(* IEC 61131-3 sources: JingjiangMoonbox/Application/Application/任务列表/Main_Task/IO列表 (part 2) *)

(* ---- KS_FB_MapAxisIOExtra.st ---- *)
(*@CES
Name=KS_FB_MapAxisIOExtra
Type=FunctionBlock
TypeGuid=6f9dac99-8de1-4efc-8465-68ac443b7d08
Guid=6be90e54-b934-4bee-925a-ddca26256504
HasDeclaration=True
HasImplementation=True
*)
{DECLARATION}
FUNCTION_BLOCK KS_FB_MapAxisIOExtra
VAR_INPUT
	i_xEn									: BOOL;(*功能块使能|*)
	i_xEnableInput							: BOOL;(*使能输入|*)
	i_xEnableOutput							: BOOL;(*使能输出|*)
	i_pstStIOMap_Axis_Extra_FE			: POINTER TO StIOMap_Axis_Extra_FE;(*轴io数据区域|*)

	i_xPreHeating							: BOOL; (* 预加热 *)
	i_xPreHeating_Err						: BOOL; (* 预加热报警\温控信号 *)
	i_xPreHotBlower							: BOOL; (* 预热风 *)
	i_xPreHotBlower_Err						: BOOL; (* 预热风报警 *)
	i_xCoolBlower							: BOOL; (* 冷风开关 *)
	i_xCoolBlower_Button					: BOOL; (* 冷风按钮 *)
	i_xCoolBlower_Err						: BOOL; (* 冷风报警 *)
	i_xHotBlower							: BOOL; (* 热风开关 *)
	i_xHotBlower_Button						: BOOL; (* 热风按钮 *)
	i_xHotBlower_Err						: BOOL; (* 热风报警 *)
	i_xHotBlower_Opened_Act					: BOOL; (* 热风实际被打开了|2022.5.11.192858|没有反馈时候需要写true*)
	i_xHotBlower_CHNL2						: BOOL; (* 第2路热风开关 *)
	i_xHotBlower_Button_CHNL2				: BOOL; (* 第2路热风按钮 *)
	i_xHotBlower_Err_CHNL2					: BOOL; (* 第2路热风报警 *)
	i_xHotBlower_Opened_Act_CHNL2			: BOOL; (* 热风2实际被打开了|2022.5.11.192858|没有反馈时候需要写true*)
	i_xTemReachToTarget						: BOOL; (* 到达目标温度 *)
	i_xSteamHeating							: BOOL; (* 蒸汽加热开关 *)
	i_xSteamHeating_Err						: BOOL; (* 蒸汽加热报警 *)
	i_xHeating_I							: BOOL; (* 电加热I档 *)
	i_xHeating_II							: BOOL; (* 电加热II档 *)
	i_xHeating_III							: BOOL; (* 电加热III档 *)
	i_xHeating_Button						: BOOL; (* 加热按钮 *)
	i_xHeating_I_CHNL2						: BOOL; (* 第2路电加热I档 *)
	i_xHeating_II_CHNL2						: BOOL; (* 第2路电加热II档 *)
	i_xHeating_III_CHNL2					: BOOL; (* 第2路电加热III档 *)
	i_xHeating_Button_CHNL2					: BOOL; (* 第2路加热按钮 *)
	i_xAllExhBlower_Up						: BOOL; (* 全上排风 *)
	i_xAllExhBlower_Err_Up					: BOOL; (* 上排风报警 *)
	i_xAllExhBlower_Dn						: BOOL; (* 全下排风 *)
	i_xAllExhBlower_Err_Dn					: BOOL; (* 下排风报警 *)
	i_xAllCoolBlower						: BOOL; (* 全冷风 *)
	i_xAllHotBlower							: BOOL; (* 全热风 *)
	i_xAllHeating							: BOOL; (* 全加热 *)
	i_xAirInletMotorMin_Limit				: BOOL; (* 进风口风门电机最小开度限位 *)
	i_xAirInletMotorMax_Limit				: BOOL; (* 进风口风门电机最大开度限位 *)
	i_xOvensAirOutMotorMin_Limit			: BOOL; (* 烘箱出风口风门电机最小开度限位 *)
	i_xOvensAirOutMotorMax_Limit			: BOOL; (* 烘箱出风口风门电机最大开度限位 *)
	i_xAirExhaustMotorMin_Limit				: BOOL; (* 排风口风门电机最小开度限位 *)
	i_xAirExhaustMotorMax_Limit				: BOOL; (* 排风口风门电机最大开度限位 *)
	i_xAirReturnMotorMin_Limit				: BOOL; (* 回风口风门电机最小开度限位 *)
	i_xAirReturnMotorMax_Limit				: BOOL; (* 回风口风门电机最大开度限位 *)
	i_xScraperInveterError					: BOOL; (* 刮刀变频器报警 *)
	i_xScraperOn							: BOOL; (* 刮刀开关 *)
	i_xInkRollerInveterError				: BOOL; (* 递墨辊变频器报警 |2022.3.26.094940*)
	i_xInkRoller_CW							: BOOL; (* 递墨辊正转开 *)
	i_xInkRoller_CCW						: BOOL; (* 递墨辊反转开 *)
	i_xInkRoller_Up							: BOOL; (* 递墨辊上 *)
	i_xInkRoller_Dn							: BOOL; (* 递墨辊下 *)
	i_xTurnoverFilmAgency					: BOOL; (* 翻料架开关 *)
	i_wAI_AirInletMotor						: WORD; (* 进风口反馈|模拟量控制风门LEL *)
	i_wAI_OvensAirOutMotor					: WORD; (* 烘箱出风口反馈|模拟量控制风门LEL *)
	i_wAI_AirExhaustMotor					: WORD; (* 排风口反馈|模拟量控制风门LEL *)
	i_wAI_AirReturnMotor					: WORD; (* 回风反馈|模拟量控制风门LEL *)
	i_wInputLel								: WORD; (* LEL浓度反馈 *)
	i_wInAllAir								: WORD; (* 总进风反馈输入 *)
	i_wInFreshAir							: WORD; (* 新风反馈输入 *)
	i_wInExhaustAir							: WORD; (* 排风反馈输入 *)
	i_wInReturnAir							: WORD; (* 二次回风反馈输入 *)
	i_xTaper_Incr							: BOOL; (* 增加锥度+|针对牵引 *)
	i_xTaper_Decr							: BOOL; (* 减小锥度-|针对牵引 *)
	i_wAI_CoatingSensor						: WORD; (* 涂布传感器模拟量 *)
	i_byAIType_CoatingSensor				: BYTE; (* 涂布传感器类型 *)
	i_xAirExhaustSwitch						: BOOL; (* 色组排风输入开关 *)
	i_xAirExhaustButton						: BOOL; (* 色组排风输入按钮 *)
	i_xPushIn_PrnRoller						: BOOL; (* 顶版-进 *)
	i_xPullOut_PrnRoller					: BOOL; (* 顶版-退 *)
	i_xRsvd_DI0								: BOOL; (* 数字量输入保留0 *)
	i_xRsvd_DI1								: BOOL; (* 数字量输入保留1 *)
	i_xRsvd_DI2								: BOOL; (* 数字量输入保留2 *)
	i_xRsvd_DI3								: BOOL; (* 数字量输入保留3 *)
	i_xRsvd_DI4								: BOOL; (* 数字量输入保留4 *)
	i_xRsvd_DI5								: BOOL; (* 数字量输入保留5 *)
	i_xRsvd_DI6								: BOOL; (* 数字量输入保留6 *)
	i_xRsvd_DI7								: BOOL; (* 数字量输入保留7 *)
	i_xRsvd_DI8								: BOOL; (* 数字量输入保留8 *)
	i_xRsvd_DI9								: BOOL; (* 数字量输入保留9 *)
	i_xRsvd_DI10							: BOOL; (* 数字量输入保留10 *)
	i_xRsvd_DI11							: BOOL; (* 数字量输入保留11 *)
	i_xRsvd_DI12							: BOOL; (* 数字量输入保留12 *)
	i_xRsvd_DI13							: BOOL; (* 数字量输入保留13 *)
	i_xRsvd_DI14							: BOOL; (* 数字量输入保留14 *)
	i_xRsvd_DI15							: BOOL; (* 数字量输入保留15 *)
	i_wRsvd_AI0								: WORD; (* 模拟量输入保留0 *)
	i_wRsvd_AI1								: WORD; (* 模拟量输入保留1 *)
	i_wRsvd_AI2								: WORD; (* 模拟量输入保留2 *)
	i_wRsvd_AI3								: WORD; (* 模拟量输入保留3 *)
	i_wRsvd_AI4								: WORD; (* 模拟量输入保留4 *)
	i_wRsvd_AI5								: WORD; (* 模拟量输入保留5 *)

END_VAR
VAR_OUTPUT
	o_xEno									: BOOL;
	o_iErNo									: INT;

	o_xRel_PreHeating						: BOOL; (* 预加热接触器 *)
	o_xLamp_PreHeating						: BOOL; (* 预加热指示灯 *)
	o_xRel_ResetErr_PreHeating				: BOOL; (* 预加热故障复位 *)
	o_wAO_PreHeating						: WORD; (* 预加热模拟量 *)
	o_xRel_PreHeatingRoller_Motor			: BOOL; (* 预热辊使能 *)
	o_xRel_PreHeatingRoller_Motor_Rev		: BOOL; (* 预热辊反转使能 *)
	o_wAO_PreHeatingRoller_Motor			: WORD; (* 预热辊模拟量输出 *)
	o_xRel_PreHotBlower						: BOOL; (* 预热风接触器 *)
	o_xLamp_PreHotBlower					: BOOL; (* 预热风指示灯 *)
	o_xRel_ResetErr_PreHotBlower			: BOOL; (* 预热风故障复位 *)
	o_wAO_PreHotBlower						: WORD; (* 预热风模拟量 *)
	o_xRel_CoolBlower						: BOOL; (* 冷风接触器 *)
	o_xLamp_CoolBlower						: BOOL; (* 冷风指示灯 *)
	o_xRel_HotBlower						: BOOL; (* 热风接触器 *)
	o_xLamp_HotBlower						: BOOL; (* 热风指示灯 *)
	o_xRel_ResetErr_HotBlower				: BOOL; (* 热风故障复位 *)
	o_wAO_HotBlower							: WORD; (* 热风模拟量输出 *)
	o_xRel_HotBlower_CHNL2					: BOOL; (* 第2路热风接触器 *)
	o_xLamp_HotBlower_CHNL2					: BOOL; (* 第2路热风指示灯 *)
	o_xRel_ResetErr_HotBlower_CHNL2			: BOOL; (* 第2路热风故障复位 *)
	o_wAO_HotBlower_CHNL2					: WORD; (* 第2路热风模拟量输出 *)
	o_xRel_SteamHeating						: BOOL; (* 蒸汽输出 *)
	o_xLamp_SteamHeating					: BOOL; (* 蒸汽加热指示灯 *)
	o_xRel_ResetErr_SteamHeating			: BOOL; (* 蒸汽加热复位 *)
	o_wAO_SteamHeating						: WORD; (* 蒸汽加热模拟量输出 *)
	o_xRel_Heating_I						: BOOL; (* 电加热I档 *)
	o_xRel_Heating_II						: BOOL; (* 电加热II档 *)
	o_xRel_Heating_III						: BOOL; (* 电加热III档 *)
	o_xLamp_Heating							: BOOL; (* 电加热指示灯 *)
	o_xRel_Heating_I_CHNL2					: BOOL; (* 第2路电加热I档 *)
	o_xRel_Heating_II_CHNL2					: BOOL; (* 第2路电加热II档 *)
	o_xRel_Heating_III_CHNL2				: BOOL; (* 第2路电加热III档 *)
	o_xLamp_Heating_CHNL2					: BOOL; (* 第2路电加热指示灯 *)
	o_xRel_AllExhBlower_Up					: BOOL; (* 上排风继电器输出 *)
	o_xLamp_AllExhBlower_Up					: BOOL; (* 全上排风指示灯 *)
	o_xRel_ModeStar_AllExhBlower_Up			: BOOL; (* 上排风模式-星形 *)
	o_xRel_ModeTriangle_AllExhBlower_Up		: BOOL; (* 上排风模式-三角 *)
	o_xRel_ResetErr_AllExhBlower_Up			: BOOL; (* 上排风故障复位 *)
	o_wAO_AllExhBlower_Up					: WORD; (* 上排风模拟量输出 *)
	o_xRel_AllExhBlower_Dn					: BOOL; (* 下排风继电器输出 *)
	o_xLamp_AllExhBlower_Dn					: BOOL; (* 全下排风指示灯 *)
	o_xRel_ModeStar_AllExhBlower_Dn			: BOOL; (* 下排风模式-星形 *)
	o_xRel_ModeTriangle_AllExhBlower_Dn		: BOOL; (* 下排风模式-三角 *)
	o_xRel_ResetErr_AllExhBlower_Dn			: BOOL; (* 下排风故障复位 *)
	o_wAO_AllExhBlower_Dn					: WORD; (* 下排风模拟量输出 *)
	o_xLamp_AllCoolBlower					: BOOL; (* 全冷风指示灯 *)
	o_xLamp_AllHotBlower					: BOOL; (* 全热风指示灯 *)
	o_xLamp_AllHeating						: BOOL; (* 全加热指示灯 *)
	o_xAirInletMotor_Increase				: BOOL; (* 进风口风门开度增大 *)
	o_xAirInletMotor_Decrease				: BOOL; (* 进风口风门开度减小 *)
	o_xOvensAirOutMotor_Increase			: BOOL; (* 烘箱出风口风门开度增大 *)
	o_xOvensAirOutMotor_Decrease			: BOOL; (* 烘箱出风口风门开度减小 *)
	o_xAirExhaustMotor_Increase				: BOOL; (* 排风口风门开度增大 *)
	o_xAirExhaustMotor_Decrease				: BOOL; (* 排风口风门开度减小 *)
	o_xAirReturnMotor_Increase				: BOOL; (* 回风风门开度增大 *)
	o_xAirReturnMotor_Decrease				: BOOL; (* 回风风门开度减小 *)
	o_xScraperOn							: BOOL; (* 刮刀输出 *)
	o_xScraperRst							: BOOL;(*刮刀故障复位*)
	o_wAO_Scraper							: WORD; (* 刮刀模拟量输出 *)
	o_xInkRollerOn							: BOOL; (* 递墨辊运动信号 *)
	o_xInkRollerRst							: BOOL;(*递墨辊复位2022.7.8.093223*)
	o_xRel_InkRoller_CW						: BOOL; (* 递墨辊正转 *)
	o_xRel_InkRoller_CCW					: BOOL; (* 递墨辊反转 *)
	o_wAO_InkRoller							: WORD; (* 递墨辊模拟量输出 *)
	(*2026.05.25.135151*)
	o_wAO_InkRoller_Dir						: WORD;(* 递墨辊模拟量输出@±10V *)
	o_xRel_InkRoller_Up						: BOOL; (* 递墨辊上输出 *)
	o_xRel_InkRoller_Dn						: BOOL; (* 递墨辊下输出 *)
	o_xRel_TurnoverFilmAgency				: BOOL; (* 翻料架输出 *)
	o_xRel_ColdWaterRoller_Motor			: BOOL; (* 水冷辊电机使能 *)
	o_xRel_ColdWaterRoller_Motor_Rev		: BOOL; (* 水冷辊电机反转使能 *)
	o_wAO_ColdWaterRoller_Motor				: WORD; (* 水冷辊电机模拟量输出 *)
	o_xRel_DriveAfterPrint_Motor			: BOOL; (* 印后传动辊电机使能 *)
	o_xRel_DriveAfterPrint_Motor_Rev		: BOOL; (* 印后传动辊电机反转 *)
	o_wAO_DriveAfterPrint_Motor				: WORD; (* 印后传动辊电机模拟量输出 *)
	o_wAO_AirInletMotor						: WORD; (* 进口输出|模拟量控制风门LEL *)
	o_wAO_OvensAirOutMotor					: WORD; (* 烘箱出风口输出|模拟量控制风门LEL *)
	o_wAO_AirExhaustMotor					: WORD; (* 排风口输出|模拟量控制风门LEL *)
	o_wAO_AirReturnMotor					: WORD; (* 回风输出|模拟量控制风门LEL *)
	o_wInAllAir								: WORD; (* 总进风输出 *)
	o_wInFreshAir							: WORD; (* 新风输出 *)
	o_wInExhaustAir							: WORD; (* 排风输出 *)
	o_wInReturnAir							: WORD; (* 二次回风输出 *)
	o_wPreAirHotRollTorque					: WORD; (* 预热辊转矩输出 *)
	o_wCoolWaterRollTorque					: WORD; (* 水冷辊转矩输出 *)
	o_xAirExhaustEn							: BOOL; (* 色组排风输出使能 *)
	o_xRel_PushIn_PrnRoller					: BOOL; (* 顶版-进执行 *)
	o_xRel_PullOut_PrnRoller				: BOOL; (* 顶版-退执行 *)
	o_xRel_ModeStar_HotBlower				: BOOL; (* 热风输出-星形 *)
	o_xRel_ModeTriangle_HotBlower			: BOOL; (* 热风输出-三角 *)
	o_xRel_Oven								: BOOL; (* 色组烘箱输出 *)
	o_xRsvd_DO0								: BOOL; (* 数字量输出保留0 *)
	o_xRsvd_DO1								: BOOL; (* 数字量输出保留1 *)
	o_xRsvd_DO2								: BOOL; (* 数字量输出保留2 *)
	o_xRsvd_DO3								: BOOL; (* 数字量输出保留3 *)
	o_xRsvd_DO4								: BOOL; (* 数字量输出保留4 *)
	o_xRsvd_DO5								: BOOL; (* 数字量输出保留5 *)
	o_xRsvd_DO6								: BOOL; (* 数字量输出保留6 *)
	o_xRsvd_DO7								: BOOL; (* 数字量输出保留7 *)
	o_xRsvd_DO8								: BOOL; (* 数字量输出保留8 *)
	o_xRsvd_DO9								: BOOL; (* 数字量输出保留9 *)
	o_xRsvd_DO10							: BOOL; (* 数字量输出保留10 *)
	o_xRsvd_DO11							: BOOL; (* 数字量输出保留11 *)
	o_xRsvd_DO12							: BOOL; (* 数字量输出保留12 *)
	o_xRsvd_DO13							: BOOL; (* 数字量输出保留13 *)
	o_xRsvd_DO14							: BOOL; (* 数字量输出保留14 *)
	o_xRsvd_DO15							: BOOL; (* 数字量输出保留15 *)
	o_wRsvd_AO0								: WORD; (* 模拟量输出保留0 *)
	o_wRsvd_AO1								: WORD; (* 模拟量输出保留1 *)
	o_wRsvd_AO2								: WORD; (* 模拟量输出保留2 *)
	o_wRsvd_AO3								: WORD; (* 模拟量输出保留3 *)
	o_wRsvd_AO4								: WORD; (* 模拟量输出保留4 *)
	o_wRsvd_AO5								: WORD; (* 模拟量输出保留5 *)
END_VAR
VAR
END_VAR

{IMPLEMENTATION}
o_xEno:= i_xEn;
o_iErNo:= 0;
IF i_xEn THEN
	IF i_pstStIOMap_Axis_Extra_FE<>0 THEN
		IF i_xEnableInput THEN (* 输入 *)
			i_pstStIOMap_Axis_Extra_FE^.i_xPreHeating					:= i_xPreHeating					;//		: BOOL; (* 预加热 *)
			i_pstStIOMap_Axis_Extra_FE^.i_xPreHeating_Err				:= i_xPreHeating_Err				;//		: BOOL; (* 预加热报警\温控信号 *)
			i_pstStIOMap_Axis_Extra_FE^.i_xPreHotBlower					:= i_xPreHotBlower					;//		: BOOL; (* 预热风 *)
			i_pstStIOMap_Axis_Extra_FE^.i_xPreHotBlower_Err				:= i_xPreHotBlower_Err				;//		: BOOL; (* 预热风报警 *)
			i_pstStIOMap_Axis_Extra_FE^.i_xCoolBlower					:= i_xCoolBlower					;//		: BOOL; (* 冷风开关 *)
			i_pstStIOMap_Axis_Extra_FE^.i_xCoolBlower_Button				:= i_xCoolBlower_Button				;//		: BOOL; (* 冷风按钮 *)
			i_pstStIOMap_Axis_Extra_FE^.i_xCoolBlower_Err				:= i_xCoolBlower_Err				;//		: BOOL; (* 冷风报警 *)
			i_pstStIOMap_Axis_Extra_FE^.i_xHotBlower						:= i_xHotBlower						;//		: BOOL; (* 热风开关 *)
			i_pstStIOMap_Axis_Extra_FE^.i_xHotBlower_Button				:= i_xHotBlower_Button				;//		: BOOL; (* 热风按钮 *)
			i_pstStIOMap_Axis_Extra_FE^.i_xHotBlower_Err					:= i_xHotBlower_Err					;//		: BOOL; (* 热风报警 *)
			i_pstStIOMap_Axis_Extra_FE^.i_xHotBlower_Opened_Act			:= i_xHotBlower_Opened_Act			;//		: BOOL; (* 热风实际被打开了|2022.5.11.192858|没有反馈时候需要写true*)
			i_pstStIOMap_Axis_Extra_FE^.i_xHotBlower_CHNL2				:= i_xHotBlower_CHNL2				;//		: BOOL; (* 第2路热风开关 *)
			i_pstStIOMap_Axis_Extra_FE^.i_xHotBlower_Button_CHNL2		:= i_xHotBlower_Button_CHNL2		;//		: BOOL; (* 第2路热风按钮 *)
			i_pstStIOMap_Axis_Extra_FE^.i_xHotBlower_Err_CHNL2			:= i_xHotBlower_Err_CHNL2			;//		: BOOL; (* 第2路热风报警 *)
			i_pstStIOMap_Axis_Extra_FE^.i_xHotBlower_Opened_Act_CHNL2	:= i_xHotBlower_Opened_Act_CHNL2	;//		: BOOL; (* 热风2实际被打开了|2022.5.11.192858|没有反馈时候需要写true*)
			i_pstStIOMap_Axis_Extra_FE^.i_xTemReachToTarget				:= i_xTemReachToTarget				;//		: BOOL; (* 到达目标温度 *)
			i_pstStIOMap_Axis_Extra_FE^.i_xSteamHeating					:= i_xSteamHeating					;//		: BOOL; (* 蒸汽加热开关 *)
			i_pstStIOMap_Axis_Extra_FE^.i_xSteamHeating_Err				:= i_xSteamHeating_Err				;//		: BOOL; (* 蒸汽加热报警 *)
			i_pstStIOMap_Axis_Extra_FE^.i_xHeating_I						:= i_xHeating_I						;//		: BOOL; (* 电加热I档 *)
			i_pstStIOMap_Axis_Extra_FE^.i_xHeating_II					:= i_xHeating_II					;//		: BOOL; (* 电加热II档 *)
			i_pstStIOMap_Axis_Extra_FE^.i_xHeating_III					:= i_xHeating_III					;//		: BOOL; (* 电加热III档 *)
			i_pstStIOMap_Axis_Extra_FE^.i_xHeating_Button				:= i_xHeating_Button				;//		: BOOL; (* 加热按钮 *)
			i_pstStIOMap_Axis_Extra_FE^.i_xHeating_I_CHNL2				:= i_xHeating_I_CHNL2				;//		: BOOL; (* 第2路电加热I档 *)
			i_pstStIOMap_Axis_Extra_FE^.i_xHeating_II_CHNL2				:= i_xHeating_II_CHNL2				;//		: BOOL; (* 第2路电加热II档 *)
			i_pstStIOMap_Axis_Extra_FE^.i_xHeating_III_CHNL2				:= i_xHeating_III_CHNL2				;//		: BOOL; (* 第2路电加热III档 *)
			i_pstStIOMap_Axis_Extra_FE^.i_xHeating_Button_CHNL2			:= i_xHeating_Button_CHNL2			;//		: BOOL; (* 第2路加热按钮 *)
			i_pstStIOMap_Axis_Extra_FE^.i_xAllExhBlower_Up				:= i_xAllExhBlower_Up				;//		: BOOL; (* 全上排风 *)
			i_pstStIOMap_Axis_Extra_FE^.i_xAllExhBlower_Err_Up			:= i_xAllExhBlower_Err_Up			;//		: BOOL; (* 上排风报警 *)
			i_pstStIOMap_Axis_Extra_FE^.i_xAllExhBlower_Dn				:= i_xAllExhBlower_Dn				;//		: BOOL; (* 全下排风 *)
			i_pstStIOMap_Axis_Extra_FE^.i_xAllExhBlower_Err_Dn			:= i_xAllExhBlower_Err_Dn			;//		: BOOL; (* 下排风报警 *)
			i_pstStIOMap_Axis_Extra_FE^.i_xAllCoolBlower					:= i_xAllCoolBlower					;//		: BOOL; (* 全冷风 *)
			i_pstStIOMap_Axis_Extra_FE^.i_xAllHotBlower					:= i_xAllHotBlower					;//		: BOOL; (* 全热风 *)
			i_pstStIOMap_Axis_Extra_FE^.i_xAllHeating					:= i_xAllHeating					;//		: BOOL; (* 全加热 *)
			i_pstStIOMap_Axis_Extra_FE^.i_xAirInletMotorMin_Limit		:= i_xAirInletMotorMin_Limit		;//		: BOOL; (* 进风口风门电机最小开度限位 *)
			i_pstStIOMap_Axis_Extra_FE^.i_xAirInletMotorMax_Limit		:= i_xAirInletMotorMax_Limit		;//		: BOOL; (* 进风口风门电机最大开度限位 *)
			i_pstStIOMap_Axis_Extra_FE^.i_xOvensAirOutMotorMin_Limit		:= i_xOvensAirOutMotorMin_Limit		;//		: BOOL; (* 烘箱出风口风门电机最小开度限位 *)
			i_pstStIOMap_Axis_Extra_FE^.i_xOvensAirOutMotorMax_Limit		:= i_xOvensAirOutMotorMax_Limit		;//		: BOOL; (* 烘箱出风口风门电机最大开度限位 *)
			i_pstStIOMap_Axis_Extra_FE^.i_xAirExhaustMotorMin_Limit		:= i_xAirExhaustMotorMin_Limit		;//		: BOOL; (* 排风口风门电机最小开度限位 *)
			i_pstStIOMap_Axis_Extra_FE^.i_xAirExhaustMotorMax_Limit		:= i_xAirExhaustMotorMax_Limit		;//		: BOOL; (* 排风口风门电机最大开度限位 *)
			i_pstStIOMap_Axis_Extra_FE^.i_xAirReturnMotorMin_Limit		:= i_xAirReturnMotorMin_Limit		;//		: BOOL; (* 回风口风门电机最小开度限位 *)
			i_pstStIOMap_Axis_Extra_FE^.i_xAirReturnMotorMax_Limit		:= i_xAirReturnMotorMax_Limit		;//		: BOOL; (* 回风口风门电机最大开度限位 *)
			i_pstStIOMap_Axis_Extra_FE^.i_xScraperInveterError			:= i_xScraperInveterError			;//		: BOOL; (* 刮刀变频器报警 *)
			i_pstStIOMap_Axis_Extra_FE^.i_xScraperOn						:= i_xScraperOn						;//		: BOOL; (* 刮刀开关 *)
			i_pstStIOMap_Axis_Extra_FE^.i_xInkRollerInveterError			:= i_xInkRollerInveterError			;//		: BOOL; (* 递墨辊变频器报警 |2022.3.26.094940*)
			i_pstStIOMap_Axis_Extra_FE^.i_xInkRoller_CW					:= i_xInkRoller_CW					;//		: BOOL; (* 递墨辊正转开 *)
			i_pstStIOMap_Axis_Extra_FE^.i_xInkRoller_CCW					:= i_xInkRoller_CCW					;//		: BOOL; (* 递墨辊反转开 *)
			i_pstStIOMap_Axis_Extra_FE^.i_xInkRoller_Up					:= i_xInkRoller_Up					;//		: BOOL; (* 递墨辊上 *)
			i_pstStIOMap_Axis_Extra_FE^.i_xInkRoller_Dn					:= i_xInkRoller_Dn					;//		: BOOL; (* 递墨辊下 *)
			i_pstStIOMap_Axis_Extra_FE^.i_xTurnoverFilmAgency			:= i_xTurnoverFilmAgency			;//		: BOOL; (* 翻料架开关 *)
			i_pstStIOMap_Axis_Extra_FE^.i_wAI_AirInletMotor				:= i_wAI_AirInletMotor				;//		: WORD; (* 进风口反馈|模拟量控制风门LEL *)
			i_pstStIOMap_Axis_Extra_FE^.i_wAI_OvensAirOutMotor			:= i_wAI_OvensAirOutMotor			;//		: WORD; (* 烘箱出风口反馈|模拟量控制风门LEL *)
			i_pstStIOMap_Axis_Extra_FE^.i_wAI_AirExhaustMotor			:= i_wAI_AirExhaustMotor			;//		: WORD; (* 排风口反馈|模拟量控制风门LEL *)
			i_pstStIOMap_Axis_Extra_FE^.i_wAI_AirReturnMotor				:= i_wAI_AirReturnMotor				;//		: WORD; (* 回风反馈|模拟量控制风门LEL *)
			i_pstStIOMap_Axis_Extra_FE^.i_wInputLel						:= i_wInputLel						;//		: WORD; (* LEL浓度反馈 *)
			i_pstStIOMap_Axis_Extra_FE^.i_wInAllAir						:= i_wInAllAir						;//		: WORD; (* 总进风反馈输入 *)
			i_pstStIOMap_Axis_Extra_FE^.i_wInFreshAir					:= i_wInFreshAir					;//		: WORD; (* 新风反馈输入 *)
			i_pstStIOMap_Axis_Extra_FE^.i_wInExhaustAir					:= i_wInExhaustAir					;//		: WORD; (* 排风反馈输入 *)
			i_pstStIOMap_Axis_Extra_FE^.i_wInReturnAir					:= i_wInReturnAir					;//		: WORD; (* 二次回风反馈输入 *)
			i_pstStIOMap_Axis_Extra_FE^.i_xTaper_Incr					:= i_xTaper_Incr					;//		: BOOL; (* 增加锥度+|针对牵引 *)
			i_pstStIOMap_Axis_Extra_FE^.i_xTaper_Decr					:= i_xTaper_Decr					;//		: BOOL; (* 减小锥度-|针对牵引 *)
			i_pstStIOMap_Axis_Extra_FE^.i_wAI_CoatingSensor				:= i_wAI_CoatingSensor				;//		: WORD; (* 涂布传感器模拟量 *)
			i_pstStIOMap_Axis_Extra_FE^.i_byAIType_CoatingSensor			:= i_byAIType_CoatingSensor			;//		: BYTE; (* 涂布传感器类型 *)
			i_pstStIOMap_Axis_Extra_FE^.i_xAirExhaustSwitch				:= i_xAirExhaustSwitch				;//		: BOOL; (* 色组排风输入开关 *)
			i_pstStIOMap_Axis_Extra_FE^.i_xAirExhaustButton				:= i_xAirExhaustButton				;//		: BOOL; (* 色组排风输入按钮 *)
			i_pstStIOMap_Axis_Extra_FE^.i_xPushIn_PrnRoller				:= i_xPushIn_PrnRoller				;//		: BOOL; (* 顶版-进 *)
			i_pstStIOMap_Axis_Extra_FE^.i_xPullOut_PrnRoller				:= i_xPullOut_PrnRoller				;//		: BOOL; (* 顶版-退 *)
			i_pstStIOMap_Axis_Extra_FE^.i_xRsvd_DI0						:= i_xRsvd_DI0						;//		: BOOL; (* 数字量输入保留0 *)
			i_pstStIOMap_Axis_Extra_FE^.i_xRsvd_DI1						:= i_xRsvd_DI1						;//		: BOOL; (* 数字量输入保留1 *)
			i_pstStIOMap_Axis_Extra_FE^.i_xRsvd_DI2						:= i_xRsvd_DI2						;//		: BOOL; (* 数字量输入保留2 *)
			i_pstStIOMap_Axis_Extra_FE^.i_xRsvd_DI3						:= i_xRsvd_DI3						;//		: BOOL; (* 数字量输入保留3 *)
			i_pstStIOMap_Axis_Extra_FE^.i_xRsvd_DI4						:= i_xRsvd_DI4						;//		: BOOL; (* 数字量输入保留4 *)
			i_pstStIOMap_Axis_Extra_FE^.i_xRsvd_DI5						:= i_xRsvd_DI5						;//		: BOOL; (* 数字量输入保留5 *)
			i_pstStIOMap_Axis_Extra_FE^.i_xRsvd_DI6						:= i_xRsvd_DI6						;//		: BOOL; (* 数字量输入保留6 *)
			i_pstStIOMap_Axis_Extra_FE^.i_xRsvd_DI7						:= i_xRsvd_DI7						;//		: BOOL; (* 数字量输入保留7 *)
			i_pstStIOMap_Axis_Extra_FE^.i_xRsvd_DI8						:= i_xRsvd_DI8						;//		: BOOL; (* 数字量输入保留8 *)
			i_pstStIOMap_Axis_Extra_FE^.i_xRsvd_DI9						:= i_xRsvd_DI9						;//		: BOOL; (* 数字量输入保留9 *)
			i_pstStIOMap_Axis_Extra_FE^.i_xRsvd_DI10						:= i_xRsvd_DI10						;//		: BOOL; (* 数字量输入保留10 *)
			i_pstStIOMap_Axis_Extra_FE^.i_xRsvd_DI11						:= i_xRsvd_DI11						;//		: BOOL; (* 数字量输入保留11 *)
			i_pstStIOMap_Axis_Extra_FE^.i_xRsvd_DI12						:= i_xRsvd_DI12						;//		: BOOL; (* 数字量输入保留12 *)
			i_pstStIOMap_Axis_Extra_FE^.i_xRsvd_DI13						:= i_xRsvd_DI13						;//		: BOOL; (* 数字量输入保留13 *)
			i_pstStIOMap_Axis_Extra_FE^.i_xRsvd_DI14						:= i_xRsvd_DI14						;//		: BOOL; (* 数字量输入保留14 *)
			i_pstStIOMap_Axis_Extra_FE^.i_xRsvd_DI15						:= i_xRsvd_DI15						;//		: BOOL; (* 数字量输入保留15 *)
			i_pstStIOMap_Axis_Extra_FE^.i_wRsvd_AI0						:= i_wRsvd_AI0						;//		: WORD; (* 模拟量输入保留0 *)
			i_pstStIOMap_Axis_Extra_FE^.i_wRsvd_AI1						:= i_wRsvd_AI1						;//		: WORD; (* 模拟量输入保留1 *)
			i_pstStIOMap_Axis_Extra_FE^.i_wRsvd_AI2						:= i_wRsvd_AI2						;//		: WORD; (* 模拟量输入保留2 *)
			i_pstStIOMap_Axis_Extra_FE^.i_wRsvd_AI3						:= i_wRsvd_AI3						;//		: WORD; (* 模拟量输入保留3 *)
			i_pstStIOMap_Axis_Extra_FE^.i_wRsvd_AI4						:= i_wRsvd_AI4						;//		: WORD; (* 模拟量输入保留4 *)
			i_pstStIOMap_Axis_Extra_FE^.i_wRsvd_AI5						:= i_wRsvd_AI5						;//		: WORD; (* 模拟量输入保留5 *)

		END_IF
		IF i_xEnableOutput THEN (* 输出 *)
			o_xRel_PreHeating						:= i_pstStIOMap_Axis_Extra_FE^.o_xRel_PreHeating						  ;//: BOOL; (* 预加热接触器 *)
			o_xLamp_PreHeating						:= i_pstStIOMap_Axis_Extra_FE^.o_xLamp_PreHeating					  ;//: BOOL; (* 预加热指示灯 *)
			o_xRel_ResetErr_PreHeating				:= i_pstStIOMap_Axis_Extra_FE^.o_xRel_ResetErr_PreHeating			  ;//: BOOL; (* 预加热故障复位 *)
			o_wAO_PreHeating						:= i_pstStIOMap_Axis_Extra_FE^.o_wAO_PreHeating						  ;//: WORD; (* 预加热模拟量 *)
			o_xRel_PreHeatingRoller_Motor			:= i_pstStIOMap_Axis_Extra_FE^.o_xRel_PreHeatingRoller_Motor			  ;//: BOOL; (* 预热辊使能 *)
			o_xRel_PreHeatingRoller_Motor_Rev		:= i_pstStIOMap_Axis_Extra_FE^.o_xRel_PreHeatingRoller_Motor_Rev		  ;//: BOOL; (* 预热辊反转使能 *)
			o_wAO_PreHeatingRoller_Motor			:= i_pstStIOMap_Axis_Extra_FE^.o_wAO_PreHeatingRoller_Motor			  ;//: WORD; (* 预热辊模拟量输出 *)
			o_xRel_PreHotBlower						:= i_pstStIOMap_Axis_Extra_FE^.o_xRel_PreHotBlower					  ;//: BOOL; (* 预热风接触器 *)
			o_xLamp_PreHotBlower					:= i_pstStIOMap_Axis_Extra_FE^.o_xLamp_PreHotBlower					  ;//: BOOL; (* 预热风指示灯 *)
			o_xRel_ResetErr_PreHotBlower			:= i_pstStIOMap_Axis_Extra_FE^.o_xRel_ResetErr_PreHotBlower			  ;//: BOOL; (* 预热风故障复位 *)
			o_wAO_PreHotBlower						:= i_pstStIOMap_Axis_Extra_FE^.o_wAO_PreHotBlower					  ;//: WORD; (* 预热风模拟量 *)
			o_xRel_CoolBlower						:= i_pstStIOMap_Axis_Extra_FE^.o_xRel_CoolBlower						  ;//: BOOL; (* 冷风接触器 *)
			o_xLamp_CoolBlower						:= i_pstStIOMap_Axis_Extra_FE^.o_xLamp_CoolBlower					  ;//: BOOL; (* 冷风指示灯 *)
			o_xRel_HotBlower						:= i_pstStIOMap_Axis_Extra_FE^.o_xRel_HotBlower						  ;//: BOOL; (* 热风接触器 *)
			o_xLamp_HotBlower						:= i_pstStIOMap_Axis_Extra_FE^.o_xLamp_HotBlower						  ;//: BOOL; (* 热风指示灯 *)
			o_xRel_ResetErr_HotBlower				:= i_pstStIOMap_Axis_Extra_FE^.o_xRel_ResetErr_HotBlower				  ;//: BOOL; (* 热风故障复位 *)
			o_wAO_HotBlower							:= i_pstStIOMap_Axis_Extra_FE^.o_wAO_HotBlower						  ;//: WORD; (* 热风模拟量输出 *)
			o_xRel_HotBlower_CHNL2					:= i_pstStIOMap_Axis_Extra_FE^.o_xRel_HotBlower_CHNL2				  ;//: BOOL; (* 第2路热风接触器 *)
			o_xLamp_HotBlower_CHNL2					:= i_pstStIOMap_Axis_Extra_FE^.o_xLamp_HotBlower_CHNL2				  ;//: BOOL; (* 第2路热风指示灯 *)
			o_xRel_ResetErr_HotBlower_CHNL2			:= i_pstStIOMap_Axis_Extra_FE^.o_xRel_ResetErr_HotBlower_CHNL2		  ;//: BOOL; (* 第2路热风故障复位 *)
			o_wAO_HotBlower_CHNL2					:= i_pstStIOMap_Axis_Extra_FE^.o_wAO_HotBlower_CHNL2					  ;//: WORD; (* 第2路热风模拟量输出 *)
			o_xRel_SteamHeating						:= i_pstStIOMap_Axis_Extra_FE^.o_xRel_SteamHeating					  ;//: BOOL; (* 蒸汽输出 *)
			o_xLamp_SteamHeating					:= i_pstStIOMap_Axis_Extra_FE^.o_xLamp_SteamHeating					  ;//: BOOL; (* 蒸汽加热指示灯 *)
			o_xRel_ResetErr_SteamHeating			:= i_pstStIOMap_Axis_Extra_FE^.o_xRel_ResetErr_SteamHeating			  ;//: BOOL; (* 蒸汽加热复位 *)
			o_wAO_SteamHeating						:= i_pstStIOMap_Axis_Extra_FE^.o_wAO_SteamHeating					  ;//: WORD; (* 蒸汽加热模拟量输出 *)
			o_xRel_Heating_I						:= i_pstStIOMap_Axis_Extra_FE^.o_xRel_Heating_I						  ;//: BOOL; (* 电加热I档 *)
			o_xRel_Heating_II						:= i_pstStIOMap_Axis_Extra_FE^.o_xRel_Heating_II						  ;//: BOOL; (* 电加热II档 *)
			o_xRel_Heating_III						:= i_pstStIOMap_Axis_Extra_FE^.o_xRel_Heating_III					  ;//: BOOL; (* 电加热III档 *)
			o_xLamp_Heating							:= i_pstStIOMap_Axis_Extra_FE^.o_xLamp_Heating						  ;//: BOOL; (* 电加热指示灯 *)
			o_xRel_Heating_I_CHNL2					:= i_pstStIOMap_Axis_Extra_FE^.o_xRel_Heating_I_CHNL2				  ;//: BOOL; (* 第2路电加热I档 *)
			o_xRel_Heating_II_CHNL2					:= i_pstStIOMap_Axis_Extra_FE^.o_xRel_Heating_II_CHNL2				  ;//: BOOL; (* 第2路电加热II档 *)
			o_xRel_Heating_III_CHNL2				:= i_pstStIOMap_Axis_Extra_FE^.o_xRel_Heating_III_CHNL2				  ;//: BOOL; (* 第2路电加热III档 *)
			o_xLamp_Heating_CHNL2					:= i_pstStIOMap_Axis_Extra_FE^.o_xLamp_Heating_CHNL2					  ;//: BOOL; (* 第2路电加热指示灯 *)
			o_xRel_AllExhBlower_Up					:= i_pstStIOMap_Axis_Extra_FE^.o_xRel_AllExhBlower_Up				  ;//: BOOL; (* 上排风继电器输出 *)
			o_xLamp_AllExhBlower_Up					:= i_pstStIOMap_Axis_Extra_FE^.o_xLamp_AllExhBlower_Up				  ;//: BOOL; (* 全上排风指示灯 *)
			o_xRel_ModeStar_AllExhBlower_Up			:= i_pstStIOMap_Axis_Extra_FE^.o_xRel_ModeStar_AllExhBlower_Up		  ;//: BOOL; (* 上排风模式-星形 *)
			o_xRel_ModeTriangle_AllExhBlower_Up		:= i_pstStIOMap_Axis_Extra_FE^.o_xRel_ModeTriangle_AllExhBlower_Up	  ;//: BOOL; (* 上排风模式-三角 *)
			o_xRel_ResetErr_AllExhBlower_Up			:= i_pstStIOMap_Axis_Extra_FE^.o_xRel_ResetErr_AllExhBlower_Up		  ;//: BOOL; (* 上排风故障复位 *)
			o_wAO_AllExhBlower_Up					:= i_pstStIOMap_Axis_Extra_FE^.o_wAO_AllExhBlower_Up					  ;//: WORD; (* 上排风模拟量输出 *)
			o_xRel_AllExhBlower_Dn					:= i_pstStIOMap_Axis_Extra_FE^.o_xRel_AllExhBlower_Dn				  ;//: BOOL; (* 下排风继电器输出 *)
			o_xLamp_AllExhBlower_Dn					:= i_pstStIOMap_Axis_Extra_FE^.o_xLamp_AllExhBlower_Dn				  ;//: BOOL; (* 全下排风指示灯 *)
			o_xRel_ModeStar_AllExhBlower_Dn			:= i_pstStIOMap_Axis_Extra_FE^.o_xRel_ModeStar_AllExhBlower_Dn		  ;//: BOOL; (* 下排风模式-星形 *)
			o_xRel_ModeTriangle_AllExhBlower_Dn		:= i_pstStIOMap_Axis_Extra_FE^.o_xRel_ModeTriangle_AllExhBlower_Dn	  ;//: BOOL; (* 下排风模式-三角 *)
			o_xRel_ResetErr_AllExhBlower_Dn			:= i_pstStIOMap_Axis_Extra_FE^.o_xRel_ResetErr_AllExhBlower_Dn		  ;//: BOOL; (* 下排风故障复位 *)
			o_wAO_AllExhBlower_Dn					:= i_pstStIOMap_Axis_Extra_FE^.o_wAO_AllExhBlower_Dn					  ;//: WORD; (* 下排风模拟量输出 *)
			o_xLamp_AllCoolBlower					:= i_pstStIOMap_Axis_Extra_FE^.o_xLamp_AllCoolBlower					  ;//: BOOL; (* 全冷风指示灯 *)
			o_xLamp_AllHotBlower					:= i_pstStIOMap_Axis_Extra_FE^.o_xLamp_AllHotBlower					  ;//: BOOL; (* 全热风指示灯 *)
			o_xLamp_AllHeating						:= i_pstStIOMap_Axis_Extra_FE^.o_xLamp_AllHeating					  ;//: BOOL; (* 全加热指示灯 *)
			o_xAirInletMotor_Increase				:= i_pstStIOMap_Axis_Extra_FE^.o_xAirInletMotor_Increase				  ;//: BOOL; (* 进风口风门开度增大 *)
			o_xAirInletMotor_Decrease				:= i_pstStIOMap_Axis_Extra_FE^.o_xAirInletMotor_Decrease				  ;//: BOOL; (* 进风口风门开度减小 *)
			o_xOvensAirOutMotor_Increase			:= i_pstStIOMap_Axis_Extra_FE^.o_xOvensAirOutMotor_Increase			  ;//: BOOL; (* 烘箱出风口风门开度增大 *)
			o_xOvensAirOutMotor_Decrease			:= i_pstStIOMap_Axis_Extra_FE^.o_xOvensAirOutMotor_Decrease			  ;//: BOOL; (* 烘箱出风口风门开度减小 *)
			o_xAirExhaustMotor_Increase				:= i_pstStIOMap_Axis_Extra_FE^.o_xAirExhaustMotor_Increase			  ;//: BOOL; (* 排风口风门开度增大 *)
			o_xAirExhaustMotor_Decrease				:= i_pstStIOMap_Axis_Extra_FE^.o_xAirExhaustMotor_Decrease			  ;//: BOOL; (* 排风口风门开度减小 *)
			o_xAirReturnMotor_Increase				:= i_pstStIOMap_Axis_Extra_FE^.o_xAirReturnMotor_Increase			  ;//: BOOL; (* 回风风门开度增大 *)
			o_xAirReturnMotor_Decrease				:= i_pstStIOMap_Axis_Extra_FE^.o_xAirReturnMotor_Decrease			  ;//: BOOL; (* 回风风门开度减小 *)
			o_xScraperOn							:= i_pstStIOMap_Axis_Extra_FE^.o_xScraperOn							  ;//: BOOL; (* 刮刀输出 *)
			o_xScraperRst							:= i_pstStIOMap_Axis_Extra_FE^.o_xScraperRst							  ;//: BOOL;(*刮刀故障复位*)
			o_wAO_Scraper							:= i_pstStIOMap_Axis_Extra_FE^.o_wAO_Scraper							  ;//: WORD; (* 刮刀模拟量输出 *)
			o_xInkRollerOn							:= i_pstStIOMap_Axis_Extra_FE^.o_xInkRollerOn						  ;//: BOOL; (* 递墨辊运动信号 *)
			o_xInkRollerRst							:= i_pstStIOMap_Axis_Extra_FE^.o_xInkRollerRst						  ;//: BOOL;(*递墨辊复位2022.7.8.093223*)
			o_xRel_InkRoller_CW						:= i_pstStIOMap_Axis_Extra_FE^.o_xRel_InkRoller_CW					  ;//: BOOL; (* 递墨辊正转 *)
			o_xRel_InkRoller_CCW					:= i_pstStIOMap_Axis_Extra_FE^.o_xRel_InkRoller_CCW					  ;//: BOOL; (* 递墨辊反转 *)
			o_wAO_InkRoller							:= i_pstStIOMap_Axis_Extra_FE^.o_wAO_InkRoller						  ;//: WORD; (* 递墨辊模拟量输出 *)
			//2026.05.25.134954
			o_wAO_InkRoller_Dir						:= i_pstStIOMap_Axis_Extra_FE^.o_wAO_InkRoller_Dir				 	 ;//: WORD; (* 递墨辊模拟量输出@±10V *)
			o_xRel_InkRoller_Up						:= i_pstStIOMap_Axis_Extra_FE^.o_xRel_InkRoller_Up					  ;//: BOOL; (* 递墨辊上输出 *)
			o_xRel_InkRoller_Dn						:= i_pstStIOMap_Axis_Extra_FE^.o_xRel_InkRoller_Dn					  ;//: BOOL; (* 递墨辊下输出 *)
			o_xRel_TurnoverFilmAgency				:= i_pstStIOMap_Axis_Extra_FE^.o_xRel_TurnoverFilmAgency				  ;//: BOOL; (* 翻料架输出 *)
			o_xRel_ColdWaterRoller_Motor			:= i_pstStIOMap_Axis_Extra_FE^.o_xRel_ColdWaterRoller_Motor			  ;//: BOOL; (* 水冷辊电机使能 *)
			o_xRel_ColdWaterRoller_Motor_Rev		:= i_pstStIOMap_Axis_Extra_FE^.o_xRel_ColdWaterRoller_Motor_Rev		  ;//: BOOL; (* 水冷辊电机反转使能 *)
			o_wAO_ColdWaterRoller_Motor				:= i_pstStIOMap_Axis_Extra_FE^.o_wAO_ColdWaterRoller_Motor			  ;//: WORD; (* 水冷辊电机模拟量输出 *)
			o_xRel_DriveAfterPrint_Motor			:= i_pstStIOMap_Axis_Extra_FE^.o_xRel_DriveAfterPrint_Motor			  ;//: BOOL; (* 印后传动辊电机使能 *)
			o_xRel_DriveAfterPrint_Motor_Rev		:= i_pstStIOMap_Axis_Extra_FE^.o_xRel_DriveAfterPrint_Motor_Rev		  ;//: BOOL; (* 印后传动辊电机反转 *)
			o_wAO_DriveAfterPrint_Motor				:= i_pstStIOMap_Axis_Extra_FE^.o_wAO_DriveAfterPrint_Motor			  ;//: WORD; (* 印后传动辊电机模拟量输出 *)
			o_wAO_AirInletMotor						:= i_pstStIOMap_Axis_Extra_FE^.o_wAO_AirInletMotor					  ;//: WORD; (* 进口输出|模拟量控制风门LEL *)
			o_wAO_OvensAirOutMotor					:= i_pstStIOMap_Axis_Extra_FE^.o_wAO_OvensAirOutMotor				  ;//: WORD; (* 烘箱出风口输出|模拟量控制风门LEL *)
			o_wAO_AirExhaustMotor					:= i_pstStIOMap_Axis_Extra_FE^.o_wAO_AirExhaustMotor					  ;//: WORD; (* 排风口输出|模拟量控制风门LEL *)
			o_wAO_AirReturnMotor					:= i_pstStIOMap_Axis_Extra_FE^.o_wAO_AirReturnMotor					  ;//: WORD; (* 回风输出|模拟量控制风门LEL *)
			o_wInAllAir								:= i_pstStIOMap_Axis_Extra_FE^.o_wInAllAir							  ;//: WORD; (* 总进风输出 *)
			o_wInFreshAir							:= i_pstStIOMap_Axis_Extra_FE^.o_wInFreshAir							  ;//: WORD; (* 新风输出 *)
			o_wInExhaustAir							:= i_pstStIOMap_Axis_Extra_FE^.o_wInExhaustAir						  ;//: WORD; (* 排风输出 *)
			o_wInReturnAir							:= i_pstStIOMap_Axis_Extra_FE^.o_wInReturnAir						  ;//: WORD; (* 二次回风输出 *)
			o_wPreAirHotRollTorque					:= i_pstStIOMap_Axis_Extra_FE^.o_wPreAirHotRollTorque				  ;//: WORD; (* 预热辊转矩输出 *)
			o_wCoolWaterRollTorque					:= i_pstStIOMap_Axis_Extra_FE^.o_wCoolWaterRollTorque				  ;//: WORD; (* 水冷辊转矩输出 *)
			o_xAirExhaustEn							:= i_pstStIOMap_Axis_Extra_FE^.o_xAirExhaustEn						  ;//: BOOL; (* 色组排风输出使能 *)
			o_xRel_PushIn_PrnRoller					:= i_pstStIOMap_Axis_Extra_FE^.o_xRel_PushIn_PrnRoller				  ;//: BOOL; (* 顶版-进执行 *)
			o_xRel_PullOut_PrnRoller				:= i_pstStIOMap_Axis_Extra_FE^.o_xRel_PullOut_PrnRoller				  ;//: BOOL; (* 顶版-退执行 *)
			o_xRel_ModeStar_HotBlower				:= i_pstStIOMap_Axis_Extra_FE^.o_xRel_ModeStar_HotBlower				  ;//: BOOL; (* 热风输出-星形 *)
			o_xRel_ModeTriangle_HotBlower			:= i_pstStIOMap_Axis_Extra_FE^.o_xRel_ModeTriangle_HotBlower			  ;//: BOOL; (* 热风输出-三角 *)
			o_xRel_Oven								:= i_pstStIOMap_Axis_Extra_FE^.o_xRel_Oven							  ;//: BOOL; (* 色组烘箱输出 *)
			o_xRsvd_DO0								:= i_pstStIOMap_Axis_Extra_FE^.o_xRsvd_DO0							  ;//: BOOL; (* 数字量输出保留0 *)
			o_xRsvd_DO1								:= i_pstStIOMap_Axis_Extra_FE^.o_xRsvd_DO1							  ;//: BOOL; (* 数字量输出保留1 *)
			o_xRsvd_DO2								:= i_pstStIOMap_Axis_Extra_FE^.o_xRsvd_DO2							  ;//: BOOL; (* 数字量输出保留2 *)
			o_xRsvd_DO3								:= i_pstStIOMap_Axis_Extra_FE^.o_xRsvd_DO3							  ;//: BOOL; (* 数字量输出保留3 *)
			o_xRsvd_DO4								:= i_pstStIOMap_Axis_Extra_FE^.o_xRsvd_DO4							  ;//: BOOL; (* 数字量输出保留4 *)
			o_xRsvd_DO5								:= i_pstStIOMap_Axis_Extra_FE^.o_xRsvd_DO5							  ;//: BOOL; (* 数字量输出保留5 *)
			o_xRsvd_DO6								:= i_pstStIOMap_Axis_Extra_FE^.o_xRsvd_DO6							  ;//: BOOL; (* 数字量输出保留6 *)
			o_xRsvd_DO7								:= i_pstStIOMap_Axis_Extra_FE^.o_xRsvd_DO7							  ;//: BOOL; (* 数字量输出保留7 *)
			o_xRsvd_DO8								:= i_pstStIOMap_Axis_Extra_FE^.o_xRsvd_DO8							  ;//: BOOL; (* 数字量输出保留8 *)
			o_xRsvd_DO9								:= i_pstStIOMap_Axis_Extra_FE^.o_xRsvd_DO9							  ;//: BOOL; (* 数字量输出保留9 *)
			o_xRsvd_DO10							:= i_pstStIOMap_Axis_Extra_FE^.o_xRsvd_DO10							  ;//: BOOL; (* 数字量输出保留10 *)
			o_xRsvd_DO11							:= i_pstStIOMap_Axis_Extra_FE^.o_xRsvd_DO11							  ;//: BOOL; (* 数字量输出保留11 *)
			o_xRsvd_DO12							:= i_pstStIOMap_Axis_Extra_FE^.o_xRsvd_DO12							  ;//: BOOL; (* 数字量输出保留12 *)
			o_xRsvd_DO13							:= i_pstStIOMap_Axis_Extra_FE^.o_xRsvd_DO13							  ;//: BOOL; (* 数字量输出保留13 *)
			o_xRsvd_DO14							:= i_pstStIOMap_Axis_Extra_FE^.o_xRsvd_DO14							  ;//: BOOL; (* 数字量输出保留14 *)
			o_xRsvd_DO15							:= i_pstStIOMap_Axis_Extra_FE^.o_xRsvd_DO15							  ;//: BOOL; (* 数字量输出保留15 *)
			o_wRsvd_AO0								:= i_pstStIOMap_Axis_Extra_FE^.o_wRsvd_AO0							  ;//: WORD; (* 模拟量输出保留0 *)
			o_wRsvd_AO1								:= i_pstStIOMap_Axis_Extra_FE^.o_wRsvd_AO1							  ;//: WORD; (* 模拟量输出保留1 *)
			o_wRsvd_AO2								:= i_pstStIOMap_Axis_Extra_FE^.o_wRsvd_AO2							  ;//: WORD; (* 模拟量输出保留2 *)
			o_wRsvd_AO3								:= i_pstStIOMap_Axis_Extra_FE^.o_wRsvd_AO3							  ;//: WORD; (* 模拟量输出保留3 *)
			o_wRsvd_AO4								:= i_pstStIOMap_Axis_Extra_FE^.o_wRsvd_AO4							  ;//: WORD; (* 模拟量输出保留4 *)
			o_wRsvd_AO5								:= i_pstStIOMap_Axis_Extra_FE^.o_wRsvd_AO5							  ;//: WORD; (* 模拟量输出保留5 *)
		END_IF
	ELSE
		o_iErNo:= -1;
	END_IF
ELSE
	o_xRel_PreHeating						:= FALSE;//: BOOL; (* 预加热接触器 *)
	o_xLamp_PreHeating						:= FALSE;//: BOOL; (* 预加热指示灯 *)
	o_xRel_ResetErr_PreHeating				:= FALSE;//: BOOL; (* 预加热故障复位 *)
	o_wAO_PreHeating						:= 0;//: WORD; (* 预加热模拟量 *)
	o_xRel_PreHeatingRoller_Motor			:= FALSE;//: BOOL; (* 预热辊使能 *)
	o_xRel_PreHeatingRoller_Motor_Rev		:= FALSE;//: BOOL; (* 预热辊反转使能 *)
	o_wAO_PreHeatingRoller_Motor			:= 0;//: WORD; (* 预热辊模拟量输出 *)
	o_xRel_PreHotBlower						:= FALSE;//: BOOL; (* 预热风接触器 *)
	o_xLamp_PreHotBlower					:= FALSE;//: BOOL; (* 预热风指示灯 *)
	o_xRel_ResetErr_PreHotBlower			:= FALSE;//: BOOL; (* 预热风故障复位 *)
	o_wAO_PreHotBlower						:= 0;//: WORD; (* 预热风模拟量 *)
	o_xRel_CoolBlower						:= FALSE;//: BOOL; (* 冷风接触器 *)
	o_xLamp_CoolBlower						:= FALSE;//: BOOL; (* 冷风指示灯 *)
	o_xRel_HotBlower						:= FALSE;//: BOOL; (* 热风接触器 *)
	o_xLamp_HotBlower						:= FALSE;//: BOOL; (* 热风指示灯 *)
	o_xRel_ResetErr_HotBlower				:= FALSE;//: BOOL; (* 热风故障复位 *)
	o_wAO_HotBlower							:= 0;//: WORD; (* 热风模拟量输出 *)
	o_xRel_HotBlower_CHNL2					:= FALSE;//: BOOL; (* 第2路热风接触器 *)
	o_xLamp_HotBlower_CHNL2					:= FALSE;//: BOOL; (* 第2路热风指示灯 *)
	o_xRel_ResetErr_HotBlower_CHNL2			:= FALSE;//: BOOL; (* 第2路热风故障复位 *)
	o_wAO_HotBlower_CHNL2					:= 0;//: WORD; (* 第2路热风模拟量输出 *)
	o_xRel_SteamHeating						:= FALSE;//: BOOL; (* 蒸汽输出 *)
	o_xLamp_SteamHeating					:= FALSE;//: BOOL; (* 蒸汽加热指示灯 *)
	o_xRel_ResetErr_SteamHeating			:= FALSE;//: BOOL; (* 蒸汽加热复位 *)
	o_wAO_SteamHeating						:= 0;//: WORD; (* 蒸汽加热模拟量输出 *)
	o_xRel_Heating_I						:= FALSE;//: BOOL; (* 电加热I档 *)
	o_xRel_Heating_II						:= FALSE;//: BOOL; (* 电加热II档 *)
	o_xRel_Heating_III						:= FALSE;//: BOOL; (* 电加热III档 *)
	o_xLamp_Heating							:= FALSE;//: BOOL; (* 电加热指示灯 *)
	o_xRel_Heating_I_CHNL2					:= FALSE;//: BOOL; (* 第2路电加热I档 *)
	o_xRel_Heating_II_CHNL2					:= FALSE;//: BOOL; (* 第2路电加热II档 *)
	o_xRel_Heating_III_CHNL2				:= FALSE;//: BOOL; (* 第2路电加热III档 *)
	o_xLamp_Heating_CHNL2					:= FALSE;//: BOOL; (* 第2路电加热指示灯 *)
	o_xRel_AllExhBlower_Up					:= FALSE;//: BOOL; (* 上排风继电器输出 *)
	o_xLamp_AllExhBlower_Up					:= FALSE;//: BOOL; (* 全上排风指示灯 *)
	o_xRel_ModeStar_AllExhBlower_Up			:= FALSE;//: BOOL; (* 上排风模式-星形 *)
	o_xRel_ModeTriangle_AllExhBlower_Up		:= FALSE;//: BOOL; (* 上排风模式-三角 *)
	o_xRel_ResetErr_AllExhBlower_Up			:= FALSE;//: BOOL; (* 上排风故障复位 *)
	o_wAO_AllExhBlower_Up					:= 0;//: WORD; (* 上排风模拟量输出 *)
	o_xRel_AllExhBlower_Dn					:= FALSE;//: BOOL; (* 下排风继电器输出 *)
	o_xLamp_AllExhBlower_Dn					:= FALSE;//: BOOL; (* 全下排风指示灯 *)
	o_xRel_ModeStar_AllExhBlower_Dn			:= FALSE;//: BOOL; (* 下排风模式-星形 *)
	o_xRel_ModeTriangle_AllExhBlower_Dn		:= FALSE;//: BOOL; (* 下排风模式-三角 *)
	o_xRel_ResetErr_AllExhBlower_Dn			:= FALSE;//: BOOL; (* 下排风故障复位 *)
	o_wAO_AllExhBlower_Dn					:= 0;//: WORD; (* 下排风模拟量输出 *)
	o_xLamp_AllCoolBlower					:= FALSE;//: BOOL; (* 全冷风指示灯 *)
	o_xLamp_AllHotBlower					:= FALSE;//: BOOL; (* 全热风指示灯 *)
	o_xLamp_AllHeating						:= FALSE;//: BOOL; (* 全加热指示灯 *)
	o_xAirInletMotor_Increase				:= FALSE;//: BOOL; (* 进风口风门开度增大 *)
	o_xAirInletMotor_Decrease				:= FALSE;//: BOOL; (* 进风口风门开度减小 *)
	o_xOvensAirOutMotor_Increase			:= FALSE;//: BOOL; (* 烘箱出风口风门开度增大 *)
	o_xOvensAirOutMotor_Decrease			:= FALSE;//: BOOL; (* 烘箱出风口风门开度减小 *)
	o_xAirExhaustMotor_Increase				:= FALSE;//: BOOL; (* 排风口风门开度增大 *)
	o_xAirExhaustMotor_Decrease				:= FALSE;//: BOOL; (* 排风口风门开度减小 *)
	o_xAirReturnMotor_Increase				:= FALSE;//: BOOL; (* 回风风门开度增大 *)
	o_xAirReturnMotor_Decrease				:= FALSE;//: BOOL; (* 回风风门开度减小 *)
	o_xScraperOn							:= FALSE;//: BOOL; (* 刮刀输出 *)
	o_xScraperRst							:= FALSE;//: BOOL;(*刮刀故障复位*)
	o_wAO_Scraper							:= 0;//: WORD; (* 刮刀模拟量输出 *)
	o_xInkRollerOn							:= FALSE;//: BOOL; (* 递墨辊运动信号 *)
	o_xInkRollerRst							:= FALSE;//: BOOL;(*递墨辊复位2022.7.8.093223*)
	o_xRel_InkRoller_CW						:= FALSE;//: BOOL; (* 递墨辊正转 *)
	o_xRel_InkRoller_CCW					:= FALSE;//: BOOL; (* 递墨辊反转 *)
	o_wAO_InkRoller							:= 0;//: WORD; (* 递墨辊模拟量输出 *)
	o_xRel_InkRoller_Up						:= FALSE;//: BOOL; (* 递墨辊上输出 *)
	o_xRel_InkRoller_Dn						:= FALSE;//: BOOL; (* 递墨辊下输出 *)
	o_xRel_TurnoverFilmAgency				:= FALSE;//: BOOL; (* 翻料架输出 *)
	o_xRel_ColdWaterRoller_Motor			:= FALSE;//: BOOL; (* 水冷辊电机使能 *)
	o_xRel_ColdWaterRoller_Motor_Rev		:= FALSE;//: BOOL; (* 水冷辊电机反转使能 *)
	o_wAO_ColdWaterRoller_Motor				:= 0;//: WORD; (* 水冷辊电机模拟量输出 *)
	o_xRel_DriveAfterPrint_Motor			:= FALSE;//: BOOL; (* 印后传动辊电机使能 *)
	o_xRel_DriveAfterPrint_Motor_Rev		:= FALSE;//: BOOL; (* 印后传动辊电机反转 *)
	o_wAO_DriveAfterPrint_Motor				:= 0;//: WORD; (* 印后传动辊电机模拟量输出 *)
	o_wAO_AirInletMotor						:= 0;//: WORD; (* 进口输出|模拟量控制风门LEL *)
	o_wAO_OvensAirOutMotor					:= 0;//: WORD; (* 烘箱出风口输出|模拟量控制风门LEL *)
	o_wAO_AirExhaustMotor					:= 0;//: WORD; (* 排风口输出|模拟量控制风门LEL *)
	o_wAO_AirReturnMotor					:= 0;//: WORD; (* 回风输出|模拟量控制风门LEL *)
	o_wInAllAir								:= 0;//: WORD; (* 总进风输出 *)
	o_wInFreshAir							:= 0;//: WORD; (* 新风输出 *)
	o_wInExhaustAir							:= 0;//: WORD; (* 排风输出 *)
	o_wInReturnAir							:= 0;//: WORD; (* 二次回风输出 *)
	o_wPreAirHotRollTorque					:= 0;//: WORD; (* 预热辊转矩输出 *)
	o_wCoolWaterRollTorque					:= 0;//: WORD; (* 水冷辊转矩输出 *)
	o_xAirExhaustEn							:= FALSE;//: BOOL; (* 色组排风输出使能 *)
	o_xRel_PushIn_PrnRoller					:= FALSE;//: BOOL; (* 顶版-进执行 *)
	o_xRel_PullOut_PrnRoller				:= FALSE;//: BOOL; (* 顶版-退执行 *)
	o_xRel_ModeStar_HotBlower				:= FALSE;//: BOOL; (* 热风输出-星形 *)
	o_xRel_ModeTriangle_HotBlower			:= FALSE;//: BOOL; (* 热风输出-三角 *)
	o_xRel_Oven								:= FALSE;//: BOOL; (* 色组烘箱输出 *)
	o_xRsvd_DO0								:= FALSE;//: BOOL; (* 数字量输出保留0 *)
	o_xRsvd_DO1								:= FALSE;//: BOOL; (* 数字量输出保留1 *)
	o_xRsvd_DO2								:= FALSE;//: BOOL; (* 数字量输出保留2 *)
	o_xRsvd_DO3								:= FALSE;//: BOOL; (* 数字量输出保留3 *)
	o_xRsvd_DO4								:= FALSE;//: BOOL; (* 数字量输出保留4 *)
	o_xRsvd_DO5								:= FALSE;//: BOOL; (* 数字量输出保留5 *)
	o_xRsvd_DO6								:= FALSE;//: BOOL; (* 数字量输出保留6 *)
	o_xRsvd_DO7								:= FALSE;//: BOOL; (* 数字量输出保留7 *)
	o_xRsvd_DO8								:= FALSE;//: BOOL; (* 数字量输出保留8 *)
	o_xRsvd_DO9								:= FALSE;//: BOOL; (* 数字量输出保留9 *)
	o_xRsvd_DO10							:= FALSE;//: BOOL; (* 数字量输出保留10 *)
	o_xRsvd_DO11							:= FALSE;//: BOOL; (* 数字量输出保留11 *)
	o_xRsvd_DO12							:= FALSE;//: BOOL; (* 数字量输出保留12 *)
	o_xRsvd_DO13							:= FALSE;//: BOOL; (* 数字量输出保留13 *)
	o_xRsvd_DO14							:= FALSE;//: BOOL; (* 数字量输出保留14 *)
	o_xRsvd_DO15							:= FALSE;//: BOOL; (* 数字量输出保留15 *)
	o_wRsvd_AO0								:= 0;//: WORD; (* 模拟量输出保留0 *)
	o_wRsvd_AO1								:= 0;//: WORD; (* 模拟量输出保留1 *)
	o_wRsvd_AO2								:= 0;//: WORD; (* 模拟量输出保留2 *)
	o_wRsvd_AO3								:= 0;//: WORD; (* 模拟量输出保留3 *)
	o_wRsvd_AO4								:= 0;//: WORD; (* 模拟量输出保留4 *)
	o_wRsvd_AO5								:= 0;//: WORD; (* 模拟量输出保留5 *)
END_IF

(* ---- KS_FB_MapIO_Main.st ---- *)
(*@CES
Name=KS_FB_MapIO_Main
Type=FunctionBlock
TypeGuid=6f9dac99-8de1-4efc-8465-68ac443b7d08
Guid=8d69e06b-f6f8-423a-a44d-88632eaed767
HasDeclaration=True
HasImplementation=True
*)
{DECLARATION}
FUNCTION_BLOCK KS_FB_MapIO_Main
VAR_INPUT
	i_xEn									: BOOL;(*功能块使能|*)
	i_xEnableInput							: BOOL;(*使能输入|*)
	i_xEnableOutput							: BOOL;(*使能输出|*)
	i_pstStIOMap_Main_FE					: POINTER TO StIOMap_Main_FE;(*轴io数据区域|*)

	i_xPrestart								: BOOL; (* 预启动 *)
	i_xInk									: BOOL; (* 空转 *)
	i_xTension								: BOOL; (* 张力投入 *)
	i_xPrint								: BOOL; (* 印刷 *)
	i_xAcc									: BOOL; (* 加速 *)
	i_xDec									: BOOL; (* 减速 *)
	i_xPressAll								: BOOL; (* 全合压 *)
	i_xUnPressAll							: BOOL; (* 全离压 *)
	i_xEstop								: BOOL; (* 急停输入 *)
	i_xStop									: BOOL; (* 停机 *)
	i_xFastStop								: BOOL; (*快停*)
	i_xAlarmBell							: BOOL; (* 警报 *)
	i_xPressMode_Auto_IF					: BOOL; (* 放牵自动合压 *)
	i_xPressMode_Manu_IF					: BOOL; (* 放牵手动合压 *)
	i_xPressMode_Auto_OF					: BOOL; (* 收牵自动合压 *)
	i_xPressMode_Manu_OF					: BOOL; (* 收牵手动合压 *)
//2025.12.29.172113增加牵引变频相关变量
	i_xInverterAlarm_If						: BOOL;(*放牵变频报警输入*)
	i_xInverterAlarm_Of						: BOOL;(*收牵变频报警输入*)
	i_xInverterAlarm						: BOOL;(*牵引变频报警输入*)
	i_xInch_If								: BOOL;(*放牵单运行*)
	i_xInch_Of								: BOOL;(*收牵单运行*)

	i_xAllExhBlower_Up						: BOOL; (* 全上排风 *)
	i_xAllExhBlower_Err_Up					: BOOL; (* 上排风报警 *)
	i_xAllExhBlower_Dn						: BOOL; (* 全下排风 *)
	i_xAllExhBlower_Err_Dn					: BOOL; (* 下排风报警 *)
	i_xAllCoolBlower						: BOOL; (* 全冷风 *)
	i_xAllHotBlower							: BOOL; (* 全热风 *)
	i_xAllHeating							: BOOL; (* 全加热 *)
	(*2024.09.28.094834//增加秦华IO*)
	i_xJumpSelection						: BOOL; (* 跳板选择开关 *)
	i_xHydraulicPower						: BOOL; (* 液压站电源开关 *)
	(*2025.02.25.90543*)
	i_xPressMode_Auto_OF1							: BOOL; (* 收卷后牵引辊自动合压 *)
	i_xPressMode_Manu_OF1							: BOOL; (* 收卷后牵引辊手动合压 *)
	i_xTapPosition_Breaking					: BOOL; (* 断料档位 *)
	i_xTapPosition_UniformInk				: BOOL; (* 匀墨档位 *)

	i_xScraperOn							: BOOL; (* 刮刀开关 *)

	i_xRsvd_DI0								: BOOL; (* 数字量输入保留0 *)//超旭-点动
	i_xRsvd_DI1								: BOOL; (* 数字量输入保留1 *)
	i_xRsvd_DI2								: BOOL; (* 数字量输入保留2 *)
	i_xRsvd_DI3								: BOOL; (* 数字量输入保留3 *)
	i_xRsvd_DI4								: BOOL; (* 数字量输入保留4 *)
	i_xRsvd_DI5								: BOOL; (* 数字量输入保留5 *)
	i_xRsvd_DI6								: BOOL; (* 数字量输入保留6 *)
	i_xRsvd_DI7								: BOOL; (* 数字量输入保留7 *)
	i_xRsvd_DI8								: BOOL; (* 数字量输入保留8 *)
	i_xRsvd_DI9								: BOOL; (* 数字量输入保留9 *)
	i_wRsvd_AI0								: WORD; (* 模拟量输入保留0 *)
	i_wRsvd_AI1								: WORD; (* 模拟量输入保留1 *)
	i_wRsvd_AI2								: WORD; (* 模拟量输入保留2 *)
	i_wRsvd_AI3								: WORD; (* 模拟量输入保留3 *)
	i_wRsvd_AI4								: WORD; (* 模拟量输入保留4 *)
	i_wRsvd_AI5								: WORD; (* 模拟量输入保留5 *)

END_VAR
VAR_OUTPUT
	o_xEno									: BOOL;
	o_iErNo									: INT;
	o_xLamp_Prestart						: BOOL; (* 预启动指示 *)
	o_xLamp_Ink								: BOOL; (* 空转指示 *)
	o_xLamp_Tension							: BOOL; (* 张力投入指示 *)
	o_xLamp_Print							: BOOL; (* 印刷指示 *)
	o_xLamp_Acc								: BOOL; (* 加速指示 *)
	o_xLamp_Dec								: BOOL; (* 减速指示 *)
	o_xLamp_AllPress						: BOOL; (* 全合压指示 *)
	o_xLamp_UnPressAll						: BOOL; (* 全离压指示 *)
	o_xLamp_Estop							: BOOL; (* 急停灯输出 *)
	o_xLamp_Stop							: BOOL; (* 指示|停机 *)
	o_xRel_AlarmBell						: BOOL; (* 报警输出 *)
	o_xRel_ArcAlarm							: BOOL; (* 整机套色报警输出 *)
	o_xLamp_Press_IF						: BOOL; (* 放牵合压指示 *)
	o_xRel_Press_IF							: BOOL; (* 放牵合压输出 *)
	o_xLamp_Press_OF						: BOOL; (* 收牵合压指示 *)
	o_xRel_Press_OF							: BOOL; (* 收牵合压输出 *)
//2025.12.29.172304增加	牵引变频控制相关
	o_xCW_If								: BOOL; (* 放牵正转 *)
	o_wAO_If								: WORD; (* 放牵输出频率 *)
	o_xCW_Of								: BOOL; (* 收牵正转 *)
	o_wAO_Of								: WORD; (* 收牵输出频率 *)
	o_xAdjustEn_If							: BOOL; (* 放牵自调使能 *)
	o_wFilm_Vel_If							: WORD; (* 放牵主机速度 *)
	o_xAdjustEn_Of							: BOOL; (* 收牵自调使能 *)
	o_wFilm_Vel_Of							: WORD; (* 收牵主机速度 *)
	o_xINVERTER_RESET						: BOOL; (* (放/收)牵引变频复位 *)
	o_xInverterReset_If						: BOOL; (* 放牵变频复位 *)
	o_xInverterReset_Of						: BOOL; (* 收牵变频复位 *)

//2023.11.18.135519
	o_xRel_AllExhBlower_Up					: BOOL; (* 上排风继电器输出 *)
	o_xLamp_AllExhBlower_Up					: BOOL; (* 全上排风指示灯 *)
	o_xRel_ModeStar_AllExhBlower_Up			: BOOL; (* 上排风模式-星形 *)
	o_xRel_ModeTriangle_AllExhBlower_Up		: BOOL; (* 上排风模式-三角 *)
	o_xRel_ResetErr_AllExhBlower_Up			: BOOL; (* 上排风故障复位 *)
	o_wAO_AllExhBlower_Up					: WORD; (* 上排风模拟量输出 *)
	o_xRel_AllExhBlower_Dn					: BOOL; (* 下排风继电器输出 *)
	o_xLamp_AllExhBlower_Dn					: BOOL; (* 全下排风指示灯 *)
	o_xRel_ModeStar_AllExhBlower_Dn			: BOOL; (* 下排风模式-星形 *)
	o_xRel_ModeTriangle_AllExhBlower_Dn		: BOOL; (* 下排风模式-三角 *)
	o_xRel_ResetErr_AllExhBlower_Dn			: BOOL; (* 下排风故障复位 *)
	o_wAO_AllExhBlower_Dn					: WORD; (* 下排风模拟量输出 *)
	o_xLamp_AllCoolBlower					: BOOL; (* 全冷风指示灯 *)
	o_xLamp_AllHotBlower					: BOOL; (* 全热风指示灯 *)
	o_xLamp_AllHeating						: BOOL; (* 全加热指示灯 *)
	o_xScraperOn							: BOOL; (* 刮刀输出 *)
	o_wAO_Scraper							: WORD; (* 刮刀模拟量输出 *)

	o_xRsvd_DO0								: BOOL; (* 数字量输出保留0 *)
	o_xRsvd_DO1								: BOOL; (* 数字量输出保留1 *)
	o_xRsvd_DO2								: BOOL; (* 数字量输出保留2 *)
	o_xRsvd_DO3								: BOOL; (* 数字量输出保留3 *)
	o_xRsvd_DO4								: BOOL; (* 数字量输出保留4 *)
	o_xRsvd_DO5								: BOOL; (* 数字量输出保留5 *)
	o_xRsvd_DO6								: BOOL; (* 数字量输出保留6 *)
	o_xRsvd_DO7								: BOOL; (* 数字量输出保留7 *)
	o_xRsvd_DO8								: BOOL; (* 数字量输出保留8 *)
	o_xRsvd_DO9								: BOOL; (* 数字量输出保留9 *)
	o_wRsvd_AO0								: WORD; (* 模拟量输出保留0 *)
	o_wRsvd_AO1								: WORD; (* 模拟量输出保留1 *)
	o_wRsvd_AO2								: WORD; (* 模拟量输出保留2 *)
	o_wRsvd_AO3								: WORD; (* 模拟量输出保留3 *)
	o_wRsvd_AO4								: WORD; (* 模拟量输出保留4 *)
	o_wRsvd_AO5								: WORD; (* 模拟量输出保留5 *)
END_VAR
VAR
	xtest: BOOL;
END_VAR

{IMPLEMENTATION}
o_xEno:= i_xEn;
o_iErNo:= 0;
IF i_xEn THEN
	IF i_pstStIOMap_Main_FE<>0 THEN
		IF i_xEnableInput THEN (* 输入 *)

			i_pstStIOMap_Main_FE^.i_xPrestart					:= i_xPrestart			; (* 预启动 *)
IF i_xPrestart THEN
	xtest:= TRUE;
END_IF
			i_pstStIOMap_Main_FE^.i_xInk							:= i_xInk				; (* 空转 *)
			i_pstStIOMap_Main_FE^.i_xTension						:= i_xTension			; (* 张力投入 *)
			i_pstStIOMap_Main_FE^.i_xPrint						:= i_xPrint				; (* 印刷 *)
			i_pstStIOMap_Main_FE^.i_xAcc							:= i_xAcc				; (* 加速 *)
			i_pstStIOMap_Main_FE^.i_xDec 						:= i_xDec				; (* 减速 *)

			i_pstStIOMap_Main_FE^.i_xPressAll					:= i_xPressAll			; (* 全合压 *)
			i_pstStIOMap_Main_FE^.i_xUnPressAll					:= i_xUnPressAll		; (* 全离压 *)
			i_pstStIOMap_Main_FE^.i_xEstop						:= i_xEstop				; (* 急停输入 *)
			i_pstStIOMap_Main_FE^.i_xStop						:= i_xStop				; (* 停机 *)
			i_pstStIOMap_Main_FE^.i_xFastStop						:= i_xFastStop				; (* 快停 *)
			i_pstStIOMap_Main_FE^.i_xAlarmBell					:= i_xAlarmBell			; (* 警报 *)
			i_pstStIOMap_Main_FE^.i_xPressMode_Auto_IF			:= i_xPressMode_Auto_IF	; (* 放牵自动合压 *)
			i_pstStIOMap_Main_FE^.i_xPressMode_Manu_IF 			:= i_xPressMode_Manu_IF	; (* 放牵手动合压 *)
			i_pstStIOMap_Main_FE^.i_xPressMode_Auto_OF			:= i_xPressMode_Auto_OF	; (* 收牵自动合压 *)
			i_pstStIOMap_Main_FE^.i_xPressMode_Manu_OF			:= i_xPressMode_Manu_OF	; (* 收牵手动合压 *)
//2025.12.30.141217
			i_pstStIOMap_Main_FE^.i_xInverterAlarm_If			:= i_xInverterAlarm_If	; (* 收牵手动合压 *)
			i_pstStIOMap_Main_FE^.i_xInverterAlarm_Of			:= i_xInverterAlarm_Of	; (* 收牵手动合压 *)
			i_pstStIOMap_Main_FE^.i_xInverterAlarm			:= i_xInverterAlarm	; (* 收牵手动合压 *)
			i_pstStIOMap_Main_FE^.i_xInch_If			:= i_xInch_If	; (* 收牵手动合压 *)
			i_pstStIOMap_Main_FE^.i_xInch_Of			:= i_xInch_Of	; (* 收牵手动合压 *)

			i_pstStIOMap_Main_FE^.i_xAllExhBlower_Up				:= i_xAllExhBlower_Up;
			i_pstStIOMap_Main_FE^.i_xAllExhBlower_Err_Up			:= i_xAllExhBlower_Err_Up;
			i_pstStIOMap_Main_FE^.i_xAllExhBlower_Dn				:= i_xAllExhBlower_Dn;
			i_pstStIOMap_Main_FE^.i_xAllExhBlower_Err_Dn			:= i_xAllExhBlower_Err_Dn;
			i_pstStIOMap_Main_FE^.i_xAllCoolBlower				:= i_xAllCoolBlower;
			i_pstStIOMap_Main_FE^.i_xAllHotBlower				:= i_xAllHotBlower;
			i_pstStIOMap_Main_FE^.i_xAllHeating					:= i_xAllHeating;
			(*2024.09.28.094834//增加秦华IO*)
			i_pstStIOMap_Main_FE^.i_xJumpSelection				:= i_xJumpSelection; (* 跳板选择开关 *)
			i_pstStIOMap_Main_FE^.i_xHydraulicPower				:= i_xHydraulicPower; (* 液压站电源开关 *)
// 			(*2025.02.25.90543*)
// 			i_pstStIOMap_Main_FLEXO^.i_xPressMode_Auto_OF1			:= i_xPressMode_Auto_OF1	; (* 收卷后牵引辊自动合压 *)
// 			i_pstStIOMap_Main_FLEXO^.i_xPressMode_Manu_OF1			:= i_xPressMode_Manu_OF1	; (* 收卷后牵引辊手动合压 *)
			i_pstStIOMap_Main_FE^.i_xTapPosition_Breaking:= i_xTapPosition_Breaking;
			i_pstStIOMap_Main_FE^.i_xTapPosition_UniformInk:= i_xTapPosition_UniformInk;
			i_pstStIOMap_Main_FE^.i_xScraperOn					:= i_xScraperOn;(*刮刀总开*)
			i_pstStIOMap_Main_FE^.i_xRsvd_DI0					:= i_xRsvd_DI0; (* 数字量输入保留0 *)
			i_pstStIOMap_Main_FE^.i_xRsvd_DI1					:= i_xRsvd_DI1; (* 数字量输入保留1 *)
			i_pstStIOMap_Main_FE^.i_xRsvd_DI2					:= i_xRsvd_DI2; (* 数字量输入保留2 *)
			i_pstStIOMap_Main_FE^.i_xRsvd_DI3					:= i_xRsvd_DI3; (* 数字量输入保留3 *)
			i_pstStIOMap_Main_FE^.i_xRsvd_DI4					:= i_xRsvd_DI4; (* 数字量输入保留4 *)
			i_pstStIOMap_Main_FE^.i_xRsvd_DI5					:= i_xRsvd_DI5; (* 数字量输入保留5 *)
			i_pstStIOMap_Main_FE^.i_xRsvd_DI6					:= i_xRsvd_DI6; (* 数字量输入保留6 *)
			i_pstStIOMap_Main_FE^.i_xRsvd_DI7					:= i_xRsvd_DI7; (* 数字量输入保留7 *)
			i_pstStIOMap_Main_FE^.i_xRsvd_DI8					:= i_xRsvd_DI8; (* 数字量输入保留8 *)
			i_pstStIOMap_Main_FE^.i_xRsvd_DI9					:= i_xRsvd_DI9; (* 数字量输入保留9 *)
			i_pstStIOMap_Main_FE^.i_wRsvd_AI0					:= i_wRsvd_AI0; (* 模拟量输入保留0 *)
			i_pstStIOMap_Main_FE^.i_wRsvd_AI1					:= i_wRsvd_AI1; (* 模拟量输入保留1 *)
			i_pstStIOMap_Main_FE^.i_wRsvd_AI2					:= i_wRsvd_AI2; (* 模拟量输入保留2 *)
			i_pstStIOMap_Main_FE^.i_wRsvd_AI3					:= i_wRsvd_AI3; (* 模拟量输入保留3 *)
			i_pstStIOMap_Main_FE^.i_wRsvd_AI4					:= i_wRsvd_AI4; (* 模拟量输入保留4 *)
			i_pstStIOMap_Main_FE^.i_wRsvd_AI5					:= i_wRsvd_AI5; (* 模拟量输入保留5 *)

		END_IF

		IF i_xEnableOutput THEN (* 输出 *)
			o_xLamp_Prestart										:= i_pstStIOMap_Main_FE^.o_xLamp_Prestart		; (* 预启动指示 *)
			o_xLamp_Ink												:= i_pstStIOMap_Main_FE^.o_xLamp_Ink 			; (* 空转指示 *)
			o_xLamp_Tension											:= i_pstStIOMap_Main_FE^.o_xLamp_Tension 		; (* 张力投入指示 *)
			o_xLamp_Print											:= i_pstStIOMap_Main_FE^.o_xLamp_Print 			; (* 印刷指示 *)
			o_xLamp_Acc												:= i_pstStIOMap_Main_FE^.o_xLamp_Acc 			; (* 加速指示 *)
			o_xLamp_Dec												:= i_pstStIOMap_Main_FE^.o_xLamp_Dec 			; (* 减速指示 *)
			o_xLamp_AllPress										:= i_pstStIOMap_Main_FE^.o_xLamp_AllPress 		; (* 全合压指示 *)
			o_xLamp_UnPressAll										:= i_pstStIOMap_Main_FE^.o_xLamp_UnPressAll 		; (* 全离压指示 *)
			o_xLamp_Estop											:= i_pstStIOMap_Main_FE^.o_xLamp_Estop 			; (* 急停灯输出 *)
			o_xLamp_Stop											:= i_pstStIOMap_Main_FE^.o_xLamp_Stop 			; (* 指示|停机 *)
			o_xRel_AlarmBell										:= i_pstStIOMap_Main_FE^.o_xRel_AlarmBell 		; (* 报警输出 *)
			o_xRel_ArcAlarm											:= i_pstStIOMap_Main_FE^.o_xRel_ArcAlarm 		; (* 整机套色报警输出 *)
			o_xLamp_Press_IF										:= i_pstStIOMap_Main_FE^.o_xLamp_Press_IF 		; (* 放牵合压指示 *)
			o_xRel_Press_IF											:= i_pstStIOMap_Main_FE^.o_xRel_Press_IF 		; (* 放牵合压输出 *)
			o_xLamp_Press_OF										:= i_pstStIOMap_Main_FE^.o_xLamp_Press_OF 		; (* 收牵合压指示 *)
			o_xRel_Press_OF											:= i_pstStIOMap_Main_FE^.o_xRel_Press_OF 		; (* 收牵合压输出 *)
//2025.12.30.141312
			o_xCW_If											:= i_pstStIOMap_Main_FE^.o_xCW_If 		; (* 收牵合压输出 *)
			o_wAO_If											:= i_pstStIOMap_Main_FE^.o_wAO_If 		; (* 收牵合压输出 *)
			o_xCW_Of											:= i_pstStIOMap_Main_FE^.o_xCW_Of 		; (* 收牵合压输出 *)
			o_wAO_Of											:= i_pstStIOMap_Main_FE^.o_wAO_Of 		; (* 收牵合压输出 *)
			o_xAdjustEn_If											:= i_pstStIOMap_Main_FE^.o_xAdjustEn_If 		; (* 收牵合压输出 *)
			o_wFilm_Vel_If											:= i_pstStIOMap_Main_FE^.o_wFilm_Vel_If 		; (* 收牵合压输出 *)
			o_xAdjustEn_Of											:= i_pstStIOMap_Main_FE^.o_xAdjustEn_Of 		; (* 收牵合压输出 *)
			o_wFilm_Vel_Of											:= i_pstStIOMap_Main_FE^.o_wFilm_Vel_Of 		; (* 收牵合压输出 *)
			o_xINVERTER_RESET											:= i_pstStIOMap_Main_FE^.o_xINVERTER_RESET 		; (* 收牵合压输出 *)
			o_xInverterReset_If											:= i_pstStIOMap_Main_FE^.o_xInverterReset_If 		; (* 收牵合压输出 *)
			o_xInverterReset_Of											:= i_pstStIOMap_Main_FE^.o_xInverterReset_Of 		; (* 收牵合压输出 *)

			o_xRel_AllExhBlower_Up								:= i_pstStIOMap_Main_FE^.o_xRel_AllExhBlower_Up;
			o_xLamp_AllExhBlower_Up								:= i_pstStIOMap_Main_FE^.o_xLamp_AllExhBlower_Up;
			o_xRel_ModeStar_AllExhBlower_Up						:= i_pstStIOMap_Main_FE^.o_xRel_ModeStar_AllExhBlower_Up;
			o_xRel_ModeTriangle_AllExhBlower_Up					:= i_pstStIOMap_Main_FE^.o_xRel_ModeTriangle_AllExhBlower_Up;
			o_xRel_ResetErr_AllExhBlower_Up						:= i_pstStIOMap_Main_FE^.o_xRel_ResetErr_AllExhBlower_Up;
			o_wAO_AllExhBlower_Up								:= i_pstStIOMap_Main_FE^.o_wAO_AllExhBlower_Up;
			o_xRel_AllExhBlower_Dn								:= i_pstStIOMap_Main_FE^.o_xRel_AllExhBlower_Dn;
			o_xLamp_AllExhBlower_Dn								:= i_pstStIOMap_Main_FE^.o_xLamp_AllExhBlower_Dn;
			o_xRel_ModeStar_AllExhBlower_Dn						:= i_pstStIOMap_Main_FE^.o_xRel_ModeStar_AllExhBlower_Dn;
			o_xRel_ModeTriangle_AllExhBlower_Dn					:= i_pstStIOMap_Main_FE^.o_xRel_ModeTriangle_AllExhBlower_Dn;
			o_xRel_ResetErr_AllExhBlower_Dn						:= i_pstStIOMap_Main_FE^.o_xRel_ResetErr_AllExhBlower_Dn;
			o_wAO_AllExhBlower_Dn								:= i_pstStIOMap_Main_FE^.o_wAO_AllExhBlower_Dn;
			o_xLamp_AllCoolBlower								:= i_pstStIOMap_Main_FE^.o_xLamp_AllCoolBlower;
			o_xLamp_AllHotBlower								:= i_pstStIOMap_Main_FE^.o_xLamp_AllHotBlower;
			o_xLamp_AllHeating									:= i_pstStIOMap_Main_FE^.o_xLamp_AllHeating;
			o_xScraperOn										:= i_pstStIOMap_Main_FE^.o_xScraperOn;
			o_wAO_Scraper										:= i_pstStIOMap_Main_FE^.o_wAO_Scraper;

			o_xRsvd_DO0						:= i_pstStIOMap_Main_FE^.o_xRsvd_DO0; (* 数字量输出保留0 *) //放牵压辊离压
			o_xRsvd_DO1						:= i_pstStIOMap_Main_FE^.o_xRsvd_DO1; (* 数字量输出保留1 *)
			o_xRsvd_DO2						:= i_pstStIOMap_Main_FE^.o_xRsvd_DO2; (* 数字量输出保留2 *)
			o_xRsvd_DO3						:= i_pstStIOMap_Main_FE^.o_xRsvd_DO3; (* 数字量输出保留3 *)
			o_xRsvd_DO4						:= i_pstStIOMap_Main_FE^.o_xRsvd_DO4; (* 数字量输出保留4 *)
			o_xRsvd_DO5						:= i_pstStIOMap_Main_FE^.o_xRsvd_DO5; (* 数字量输出保留5 *)
			o_xRsvd_DO6						:= i_pstStIOMap_Main_FE^.o_xRsvd_DO6; (* 数字量输出保留6 *)
			o_xRsvd_DO7						:= i_pstStIOMap_Main_FE^.o_xRsvd_DO7; (* 数字量输出保留7 *)
			o_xRsvd_DO8						:= i_pstStIOMap_Main_FE^.o_xRsvd_DO8; (* 数字量输出保留8 *)
			o_xRsvd_DO9						:= i_pstStIOMap_Main_FE^.o_xRsvd_DO9; (* 数字量输出保留9 *)
			o_wRsvd_AO0						:= i_pstStIOMap_Main_FE^.o_wRsvd_AO0; (* 模拟量输出保留0 *)
			o_wRsvd_AO1						:= i_pstStIOMap_Main_FE^.o_wRsvd_AO1; (* 模拟量输出保留1 *)
			o_wRsvd_AO2						:= i_pstStIOMap_Main_FE^.o_wRsvd_AO2; (* 模拟量输出保留2 *)
			o_wRsvd_AO3						:= i_pstStIOMap_Main_FE^.o_wRsvd_AO3; (* 模拟量输出保留3 *)
			o_wRsvd_AO4						:= i_pstStIOMap_Main_FE^.o_wRsvd_AO4; (* 模拟量输出保留4 *)
			o_wRsvd_AO5						:= i_pstStIOMap_Main_FE^.o_wRsvd_AO5; (* 模拟量输出保留5 *)
		END_IF
	ELSE
		o_iErNo:= -1;
	END_IF
ELSE
	o_xLamp_Prestart				:= FALSE;(* 预启动指示 *)
    o_xLamp_Ink			       		:= FALSE;(* 空转指示 *)
    o_xLamp_Tension		        	:= FALSE;(* 张力投入指示 *)
    o_xLamp_Print		        	:= FALSE;(* 印刷指示 *)
    o_xLamp_Acc			        	:= FALSE;(* 加速指示 *)
    o_xLamp_Dec			        	:= FALSE;(* 减速指示 *)
    o_xLamp_AllPress	        	:= FALSE;(* 全合压指示 *)
    o_xLamp_UnPressAll	        	:= FALSE;(* 全离压指示 *)
    o_xLamp_Estop		        	:= FALSE;(* 急停灯输出 *)
    o_xLamp_Stop		        	:= FALSE;(* 指示|停机 *)
    o_xRel_AlarmBell	        	:= FALSE;(* 报警输出 *)
    o_xRel_ArcAlarm		        	:= FALSE;(* 整机套色报警输出 *)
    o_xLamp_Press_IF	        	:= FALSE;(* 放牵合压指示 *)
    o_xRel_Press_IF		        	:= FALSE;(* 放牵合压输出 *)
    o_xLamp_Press_OF	        	:= FALSE;(* 收牵合压指示 *)
    o_xRel_Press_OF		        	:= FALSE;(* 收牵合压输出 *)

	o_xRsvd_DO0						:= FALSE; (* 数字量输出保留0 *)
	o_xRsvd_DO1						:= FALSE; (* 数字量输出保留1 *)
	o_xRsvd_DO2						:= FALSE; (* 数字量输出保留2 *)
	o_xRsvd_DO3						:= FALSE; (* 数字量输出保留3 *)
	o_xRsvd_DO4						:= FALSE; (* 数字量输出保留4 *)
	o_xRsvd_DO5						:= FALSE; (* 数字量输出保留5 *)
	o_xRsvd_DO6						:= FALSE; (* 数字量输出保留6 *)
	o_xRsvd_DO7						:= FALSE; (* 数字量输出保留7 *)
	o_xRsvd_DO8						:= FALSE; (* 数字量输出保留8 *)
	o_xRsvd_DO9						:= FALSE; (* 数字量输出保留9 *)
	o_wRsvd_AO0						:= 0; (* 模拟量输出保留0 *)
	o_wRsvd_AO1						:= 0; (* 模拟量输出保留1 *)
	o_wRsvd_AO2						:= 0; (* 模拟量输出保留2 *)
	o_wRsvd_AO3						:= 0; (* 模拟量输出保留3 *)
	o_wRsvd_AO4						:= 0; (* 模拟量输出保留4 *)
	o_wRsvd_AO5						:= 0; (* 模拟量输出保留5 *)
END_IF

(* ---- KS_FB_MapIO_UwRw.st ---- *)
(*@CES
Name=KS_FB_MapIO_UwRw
Type=FunctionBlock
TypeGuid=6f9dac99-8de1-4efc-8465-68ac443b7d08
Guid=9b73f1fc-622c-41fa-a6dc-b662d2a081e6
HasDeclaration=True
HasImplementation=True
*)
{DECLARATION}
FUNCTION_BLOCK KS_FB_MapIO_UwRw
VAR_INPUT
	i_xEn									: BOOL;(*功能块使能|*)
	i_xEnableInput							: BOOL;(*使能输入|*)
	i_xEnableOutput							: BOOL;(*使能输出|*)
	i_pstStIOMap_UwRw_FE					: POINTER TO StIOMap_UwRw_FE;(*轴io数据区域|*)

	i_xEstop								: BOOL; (* 急停输入 *)
	i_xSafetyGrating						: BOOL; (* 安全光栅 *)
	i_xSafeTyGratingReset					: BOOL;	(* 安全光栅复位*)
	i_xInverterErrorA						: BOOL; (* A轴变频器故障 *)
	i_xInverterErrorB						: BOOL; (* B轴变频器故障 *)
	i_xPreCut								: BOOL; (* 预备接料 *)
	i_xCut_Cancel							: BOOL; (* 接料取消 *)
	i_xCut									: BOOL; (* 接料 *)
	i_xForward								: BOOL; (* 翻转架正转 *)
	i_xReversal								: BOOL; (* 翻转架反转 *)
	i_xAxisExchange							: BOOL; (* 轴切换 *)
	i_xIsUpCut								: BOOL; (* 上裁 *)
(*	i_xCutOnTopKnob							: BOOL; (* 上下裁 |旋钮*)*)
	i_xCutOnTopBtn							: BOOL; (* 上下裁 |按钮*)
	i_xAxisA_Locating_UpCut					: BOOL; (* 上裁A轴定位 *)
	i_xAxisB_Locating_UpCut					: BOOL; (* 上裁B轴定位 *)
	i_xAxisA_Locating_UpCut_PaperCore6Inch	: BOOL; (* 上裁A轴6寸定位 *)
	i_xAxisB_Locating_UpCut_PaperCore6Inch	: BOOL; (* 上裁B轴6寸定位 *)
(*2021.11.2.162431 替换*)
	i_xMinimumDiamProtect_UpCut				: BOOL; (* 上裁最小卷径保护 *)
	i_xAxisA_MinimumDiamProtect_UpCut		: BOOL; (* 上裁A轴最小卷径保护 *)
	i_xAxisB_MinimumDiamProtect_UpCut		: BOOL; (* 上裁B轴最小卷径保护 *)
	i_xSensor_DiamMeasureLocating_UpCut		: BOOL; (* 上裁卷径测量定位 *)
	i_xSensor_Reflex_UpCut					: BOOL; (* 上裁弧面信号 *)
	i_xAxisA_Locating_DnCut					: BOOL; (* 下裁A轴定位 *)
	i_xAxisB_Locating_DnCut					: BOOL; (* 下裁B轴定位 *)
	i_xAxisA_Locating_DnCut_PaperCore6Inch	: BOOL; (* 下裁A轴6寸定位 *)
	i_xAxisB_Locating_DnCut_PaperCore6Inch	: BOOL; (* 下裁B轴6寸定位 *)
(*2021.11.2.162446 替换*)
	i_xMinimumDiamProtect_DnCut				: BOOL; (* 下裁最小卷径保护 *)
	i_xAxisA_MinimumDiamProtect_DnCut		: BOOL; (* 下裁A轴最小卷径保护 *)
	i_xAxisB_MinimumDiamProtect_DnCut		: BOOL; (* 下裁B轴最小卷径保护 *)
	i_xSensor_DiamMeasureLocating_DnCut		: BOOL; (* 下裁卷径测量定位 *)
	i_xSensor_Reflex_DnCut					: BOOL; (* 下裁弧面信号 *)
	i_xSensor_Reflex_A_Up						: BOOL; (* A轴弧面信号 *)
	i_xSensor_Reflex_B_Up						: BOOL; (* B轴弧面信号 *)
	i_xSensor_Reflex_A_Dn						: BOOL; (* A轴弧面信号 *)
	i_xSensor_Reflex_B_Dn						: BOOL; (* B轴弧面信号 *)
	i_xPaperCoreSelect6Inch					: BOOL; (* 6寸纸管有效 *)
	i_xInverterManuReset					: BOOL; (* 变频器故障手动复位 *)
	i_xTaper_Incr							: BOOL; (* 增加锥度 *)
	i_xTaper_Decr							: BOOL; (* 减小锥度 *)
	i_xAxisInch								: BOOL; (* 轴单运行 |2022.5.24.091430*)
	(*2024.09.28.094834//增加秦华IO*)
	i_xOperation_UWRW						: BOOL; (* 收放卷运行信号 *)
	i_xSynchronous							: BOOL; (* 同步信号 *)

	i_xRsvd_DI0								: BOOL; (* 数字量输入保留0 *)
	i_xRsvd_DI1								: BOOL; (* 数字量输入保留1 *)
	i_xRsvd_DI2								: BOOL; (* 数字量输入保留2 *)
	i_xRsvd_DI3								: BOOL; (* 数字量输入保留3 *)
	i_xRsvd_DI4								: BOOL; (* 数字量输入保留4 *)
	i_xRsvd_DI5								: BOOL; (* 数字量输入保留5 *)
	i_xRsvd_DI6								: BOOL; (* 数字量输入保留6 *)
	i_xRsvd_DI7								: BOOL; (* 数字量输入保留7 *)
	i_xRsvd_DI8								: BOOL; (* 数字量输入保留8 *)
	i_xRsvd_DI9								: BOOL; (* 数字量输入保留9 *)
	i_wRsvd_AI0								: WORD; (* 模拟量输入保留0 *)
	i_wRsvd_AI1								: WORD; (* 模拟量输入保留1 *)
	i_wRsvd_AI2								: WORD; (* 模拟量输入保留2 *)
	i_wRsvd_AI3								: WORD; (* 模拟量输入保留3 *)
	i_wRsvd_AI4								: WORD; (* 模拟量输入保留4 *)
	i_wRsvd_AI5								: WORD; (* 模拟量输入保留5 *)

END_VAR
VAR_OUTPUT
	o_xEno									: BOOL;
	o_iErNo									: INT;
	o_xEstopLamp							: BOOL; (* 急停指示 *)
	o_xInverterResetA						: BOOL; (* A轴变频复位 *)
	o_xInverterResetB						: BOOL; (* B轴变频复位 *)
	o_xLamp_InverterError_A					: BOOL; (* A轴变频故障指示 *)
	o_xLamp_InverterError_B					: BOOL; (* B轴变频故障指示 *)
	o_xInverterReset_ALL					: BOOL; (* 变频器整体复位 *)
	o_xLamp_InverterError_ALL				: BOOL; (* 整机变频故障指示 *)
	o_xLamp_PreDrive						: BOOL; (* 预驱同步指示 *)
	o_xRel_TowerForeward					: BOOL; (* 塔台正转 *)
	o_xRel_TowerReversal					: BOOL; (* 塔台反转 *)
	o_xAxisALamp							: BOOL; (* A轴指示 *)
	o_xAxisBLamp							: BOOL; (* B轴指示 *)
	o_xAxisAForeward						: BOOL; (* A轴正转 *)
	o_xAxisBForeward						: BOOL; (* B轴正转 *)
	o_xCutOnTop								: BOOL; (* 上裁刀*)

	//2026.04.02.102225 | + |
	o_xCutHolder						: BOOL; (* 上裁刀架 *)
	o_xCutCylinder						: BOOL; (* 上裁胶辊 *)
	o_xCutter							: BOOL; (* 上裁裁刀 *)

	o_xCutHolder_UpCut						: BOOL; (* 上裁刀架 *)
	o_xCutCylinder_UpCut					: BOOL; (* 上裁胶辊 *)
	o_xCutter_UpCut							: BOOL; (* 上裁裁刀 *)
	o_xCutHolder_DnCut						: BOOL; (* 下裁刀架 *)
	o_xCutCylinder_DnCut					: BOOL; (* 下裁胶辊 *)
	o_xCutter_DnCut							: BOOL; (* 下裁裁刀 *)
	o_xLamp_PaperCoreSelect6Inch			: BOOL; (* 6寸纸管指示 *)
	o_xLamp_InverterError					: BOOL; (* 变频器故障指示 *)
	o_xAxisATorqueCancel					: BOOL; (* A轴转矩取消 *)
	o_xAxisBTorqueCancel					: BOOL; (* B轴转矩取消 *)
	o_wAxisATorqueVolt						: WORD; (* A轴转矩电压 *)
	o_wAxisBTorqueVolt						: WORD; (* B轴转矩电压 *)
	o_xLampAxisInching						: BOOL; (* 轴单运行中*)

	(*2024.09.28.094834//增加秦华IO*)
	o_xHydrPumpPower						: BOOL; (* 液压泵电源开关 *)
	o_xAdvanceAllBoot						: BOOL; (* 开机整体进版信号 *)
	o_xStopBack								: BOOL; (* 停止退版信号 *)
	o_xOutputAlarm							: BOOL; (* 警报输出 *)
	o_xLampInk								: BOOL; (* 空转信号 *)
	o_xServoError							: BOOL; (* 伺服故障信号 *)

	o_xRsvd_DO0								: BOOL; (* 数字量输出保留0 *)
	o_xRsvd_DO1								: BOOL; (* 数字量输出保留1 *)
	o_xRsvd_DO2								: BOOL; (* 数字量输出保留2 *)
	o_xRsvd_DO3								: BOOL; (* 数字量输出保留3 *)
	o_xRsvd_DO4								: BOOL; (* 数字量输出保留4 *)
	o_xRsvd_DO5								: BOOL; (* 数字量输出保留5 *)
	o_xRsvd_DO6								: BOOL; (* 数字量输出保留6 *)
	o_xRsvd_DO7								: BOOL; (* 数字量输出保留7 *)
	o_xRsvd_DO8								: BOOL; (* 数字量输出保留8 *)
	o_xRsvd_DO9								: BOOL; (* 数字量输出保留9 *)
	o_wRsvd_AO0								: WORD; (* 模拟量输出保留0 *)
	o_wRsvd_AO1								: WORD; (* 模拟量输出保留1 *)
	o_wRsvd_AO2								: WORD; (* 模拟量输出保留2 *)
	o_wRsvd_AO3								: WORD; (* 模拟量输出保留3 *)
	o_wRsvd_AO4								: WORD; (* 模拟量输出保留4 *)
	o_wRsvd_AO5								: WORD; (* 模拟量输出保留5 *)
END_VAR
VAR
END_VAR

{IMPLEMENTATION}
o_xEno:= i_xEn;
o_iErNo:= 0;
IF i_xEn THEN
	IF i_pstStIOMap_UwRw_FE<>0 THEN
		IF i_xEnableInput THEN (* 输入 *)

			i_pstStIOMap_UwRw_FE^.i_xEstop := i_xEstop																; (* 急停输入 *)
			i_pstStIOMap_UwRw_FE^.i_xSafetyGrating := i_xSafetyGrating												; (* 安全光栅 *)
			i_pstStIOMap_UwRw_FE^.i_xSafeTyGratingReset := i_xSafeTyGratingReset										; (* 安全光栅复位 *)
			i_pstStIOMap_UwRw_FE^.i_xInverterErrorA := i_xInverterErrorA												; (* A轴变频报警 *)
			i_pstStIOMap_UwRw_FE^.i_xInverterErrorB := i_xInverterErrorB												; (* B轴变频报警 *)
			i_pstStIOMap_UwRw_FE^.i_xPreCut := i_xPreCut																; (* 预备接料 *)
			i_pstStIOMap_UwRw_FE^.i_xCut_Cancel := i_xCut_Cancel														; (* 接料取消 *)
			i_pstStIOMap_UwRw_FE^.i_xCut := i_xCut																	; (* 接料 *)
			i_pstStIOMap_UwRw_FE^.i_xForward := i_xForward															; (* 翻转架正转 *)
			i_pstStIOMap_UwRw_FE^.i_xReversal := i_xReversal															; (* 翻转架反转 *)
			i_pstStIOMap_UwRw_FE^.i_xAxisExchange := i_xAxisExchange													; (* 轴切换 *)
			i_pstStIOMap_UwRw_FE^.i_xIsUpCut := i_xIsUpCut															; (* 上裁 |旋钮*)
			i_pstStIOMap_UwRw_FE^.i_xCutOnTopBtn := i_xCutOnTopBtn													; (* 上\下裁 |按钮*)
			i_pstStIOMap_UwRw_FE^.i_xAxisA_Locating_UpCut := i_xAxisA_Locating_UpCut									; (* 上裁A轴定位 *)
			i_pstStIOMap_UwRw_FE^.i_xAxisB_Locating_UpCut := i_xAxisB_Locating_UpCut									; (* 上裁B轴定位 *)
			i_pstStIOMap_UwRw_FE^.i_xAxisA_Locating_UpCut_PaperCore6Inch := i_xAxisA_Locating_UpCut_PaperCore6Inch	; (* 上裁A轴6寸定位 *)
			i_pstStIOMap_UwRw_FE^.i_xAxisB_Locating_UpCut_PaperCore6Inch := i_xAxisB_Locating_UpCut_PaperCore6Inch	; (* 上裁B轴6寸定位 *)

			i_pstStIOMap_UwRw_FE^.i_xMinimumDiamProtect_UpCut := i_xMinimumDiamProtect_UpCut							; (* 上裁最小卷径保护 *)

			i_pstStIOMap_UwRw_FE^.i_xAxisA_MinimumDiamProtect_UpCut := i_xAxisA_MinimumDiamProtect_UpCut				; (* 上裁A轴最小卷径保护 *)
			i_pstStIOMap_UwRw_FE^.i_xAxisB_MinimumDiamProtect_UpCut := i_xAxisB_MinimumDiamProtect_UpCut				; (* 上裁A轴最小卷径保护 *)
			i_pstStIOMap_UwRw_FE^.i_xSensor_DiamMeasureLocating_UpCut := i_xSensor_DiamMeasureLocating_UpCut			; (* 上裁卷径测量定位 *)
			i_pstStIOMap_UwRw_FE^.i_xSensor_Reflex_UpCut := i_xSensor_Reflex_UpCut								; (* 上裁弧面信号 *)
			i_pstStIOMap_UwRw_FE^.i_xAxisA_Locating_DnCut := i_xAxisA_Locating_DnCut									; (* 下裁A轴定位 *)
			i_pstStIOMap_UwRw_FE^.i_xAxisB_Locating_DnCut := i_xAxisB_Locating_DnCut									; (* 下裁B轴定位 翻转架 *)
			i_pstStIOMap_UwRw_FE^.i_xAxisA_Locating_DnCut_PaperCore6Inch := i_xAxisA_Locating_DnCut_PaperCore6Inch	; (* 下裁A轴6寸定位 *)
			i_pstStIOMap_UwRw_FE^.i_xAxisB_Locating_DnCut_PaperCore6Inch := i_xAxisB_Locating_DnCut_PaperCore6Inch	; (* 下裁B轴6寸定位 *)
			i_pstStIOMap_UwRw_FE^.i_xMinimumDiamProtect_DnCut := i_xMinimumDiamProtect_DnCut							; (* 下裁最小卷径保护 *)

			i_pstStIOMap_UwRw_FE^.i_xAxisA_MinimumDiamProtect_DnCut := i_xAxisA_MinimumDiamProtect_DnCut				; (* 下裁A轴最小卷径保护 *)
			i_pstStIOMap_UwRw_FE^.i_xAxisB_MinimumDiamProtect_DnCut := i_xAxisB_MinimumDiamProtect_DnCut				; (* 下裁A轴最小卷径保护 *)
			i_pstStIOMap_UwRw_FE^.i_xSensor_DiamMeasureLocating_DnCut := i_xSensor_DiamMeasureLocating_DnCut			; (* 下裁卷径测量定位 对射电眼 *)
			i_pstStIOMap_UwRw_FE^.i_xSensor_Reflex_DnCut := i_xSensor_Reflex_DnCut									; (* 下裁弧面信号 *)
			i_pstStIOMap_UwRw_FE^.i_xPaperCoreSelect6Inch := i_xPaperCoreSelect6Inch									; (* 6寸纸管有效 *)
			i_pstStIOMap_UwRw_FE^.i_xTaper_Incr := i_xTaper_Incr														; (* 增加锥度 *)
			i_pstStIOMap_UwRw_FE^.i_xTaper_Decr := i_xTaper_Decr														; (* 减小锥度 *)
			i_pstStIOMap_UwRw_FE^.i_xAxisInch := i_xAxisInch															; (* 轴单运行 *)
			(*2024.09.28.094834//增加秦华IO*)
			i_pstStIOMap_UwRw_FE^.i_xOperation_UWRW := i_xOperation_UWRW												; (* 收放卷运行信号 *)
			i_pstStIOMap_UwRw_FE^.i_xSynchronous := i_xSynchronous													; (* 同步信号 *)

			//2025.04.23.142158 | 弧面检测处理
			i_pstStIOMap_UwRw_FE^.i_xSensor_Reflex_A_Up := i_xSensor_Reflex_A_Up;//: BOOL; (* A轴弧面信号 *)
			i_pstStIOMap_UwRw_FE^.i_xSensor_Reflex_B_Up := i_xSensor_Reflex_B_Up;//: BOOL; (* B轴弧面信号 *)
			i_pstStIOMap_UwRw_FE^.i_xSensor_Reflex_A_Dn := i_xSensor_Reflex_A_Dn;//: BOOL; (* A轴弧面信号 *)
			i_pstStIOMap_UwRw_FE^.i_xSensor_Reflex_B_Dn := i_xSensor_Reflex_B_Dn;//: BOOL; (* B轴弧面信号 *)

			i_pstStIOMap_UwRw_FE^.i_xRsvd_DI0 := i_xRsvd_DI0															; (* 数字量输入保留0 *)//放料缺料检测
			i_pstStIOMap_UwRw_FE^.i_xRsvd_DI1 := i_xRsvd_DI1															; (* 数字量输入保留1 *)
			i_pstStIOMap_UwRw_FE^.i_xRsvd_DI2 := i_xRsvd_DI2															; (* 数字量输入保留2 *)
			i_pstStIOMap_UwRw_FE^.i_xRsvd_DI3 := i_xRsvd_DI3															; (* 数字量输入保留3 *)
			i_pstStIOMap_UwRw_FE^.i_xRsvd_DI4 := i_xRsvd_DI4															; (* 数字量输入保留4 *)
			i_pstStIOMap_UwRw_FE^.i_xRsvd_DI5 := i_xRsvd_DI5															; (* 数字量输入保留5 *)
			i_pstStIOMap_UwRw_FE^.i_xRsvd_DI6 := i_xRsvd_DI6															; (* 数字量输入保留6 *)
			i_pstStIOMap_UwRw_FE^.i_xRsvd_DI7 := i_xRsvd_DI7															; (* 数字量输入保留7 *)
			i_pstStIOMap_UwRw_FE^.i_xRsvd_DI8 := i_xRsvd_DI8															; (* 数字量输入保留8 *)
			i_pstStIOMap_UwRw_FE^.i_xRsvd_DI9 := i_xRsvd_DI9															; (* 数字量输入保留9 *)
			i_pstStIOMap_UwRw_FE^.i_wRsvd_AI0 := i_wRsvd_AI0															; (* 模拟量输入保留0 *)
			i_pstStIOMap_UwRw_FE^.i_wRsvd_AI1 := i_wRsvd_AI1															; (* 模拟量输入保留1 *)
			i_pstStIOMap_UwRw_FE^.i_wRsvd_AI2 := i_wRsvd_AI2															; (* 模拟量输入保留2 *)
			i_pstStIOMap_UwRw_FE^.i_wRsvd_AI3 := i_wRsvd_AI3															; (* 模拟量输入保留3 *)
			i_pstStIOMap_UwRw_FE^.i_wRsvd_AI4 := i_wRsvd_AI4															; (* 模拟量输入保留4 *)
			i_pstStIOMap_UwRw_FE^.i_wRsvd_AI5 := i_wRsvd_AI5															; (* 模拟量输入保留5 *)

		END_IF

		IF i_xEnableOutput THEN (* 输出 *)
			o_xEstopLamp					:= i_pstStIOMap_UwRw_FE^.o_xEstopLamp						; (* 急停指示 *)
			o_xInverterResetA				:= i_pstStIOMap_UwRw_FE^.o_xInverterResetA					; (* A轴变频复位 *)
			o_xInverterResetB				:= i_pstStIOMap_UwRw_FE^.o_xInverterResetB					; (* B轴变频复位 *)
			o_xLamp_InverterError_A				:= i_pstStIOMap_UwRw_FE^.o_xLamp_InverterError_A					; (* A轴变频故障指示 *)
			o_xLamp_InverterError_B				:= i_pstStIOMap_UwRw_FE^.o_xLamp_InverterError_B					; (* B轴变频故障指示 *)
			o_xInverterReset_ALL				:= i_pstStIOMap_UwRw_FE^.o_xInverterReset_ALL					; (* 变频故障整体复位 *)
			o_xLamp_InverterError_ALL				:= i_pstStIOMap_UwRw_FE^.o_xLamp_InverterError_ALL					; (* 整机变频故障指示 *)

			o_xLamp_PreDrive				:= i_pstStIOMap_UwRw_FE^.o_xLamp_PreDrive					; (* 预驱同步指示 *)
			o_xRel_TowerForeward			:= i_pstStIOMap_UwRw_FE^.o_xRel_TowerForeward				; (* 塔台正转 *)
			o_xRel_TowerReversal			:= i_pstStIOMap_UwRw_FE^.o_xRel_TowerReversal				; (* 塔台反转 *)
			o_xAxisALamp					:= i_pstStIOMap_UwRw_FE^.o_xAxisALamp						; (* A轴指示 *)
			o_xAxisBLamp					:= i_pstStIOMap_UwRw_FE^.o_xAxisBLamp						; (* B轴指示 *)
			o_xAxisAForeward				:= i_pstStIOMap_UwRw_FE^.o_xAxisAForeward					; (* A轴正转 *)
			o_xAxisBForeward				:= i_pstStIOMap_UwRw_FE^.o_xAxisBForeward					; (* B轴正转 *)
			o_xCutOnTop						:= i_pstStIOMap_UwRw_FE^.o_xCutOnTop							; (* 上裁刀 *)
			//2026.04.02.102225 | + |
			o_xCutHolder				:= i_pstStIOMap_UwRw_FE^.o_xCutHolder_UpCut	 OR i_pstStIOMap_UwRw_FE^.o_xCutHolder_DnCut				; (* 上裁刀架 *)
			o_xCutCylinder				:= i_pstStIOMap_UwRw_FE^.o_xCutCylinder_UpCut OR i_pstStIOMap_UwRw_FE^.o_xCutCylinder_DnCut			; (* 上裁胶辊 *)
			o_xCutter					:= i_pstStIOMap_UwRw_FE^.o_xCutter_UpCut OR i_pstStIOMap_UwRw_FE^.o_xCutter_DnCut						; (* 上裁裁刀 *)

			o_xCutHolder_UpCut				:= i_pstStIOMap_UwRw_FE^.o_xCutHolder_UpCut					; (* 上裁刀架 *)
			o_xCutCylinder_UpCut			:= i_pstStIOMap_UwRw_FE^.o_xCutCylinder_UpCut				; (* 上裁胶辊 *)
			o_xCutter_UpCut					:= i_pstStIOMap_UwRw_FE^.o_xCutter_UpCut						; (* 上裁裁刀 *)
			o_xCutHolder_DnCut				:= i_pstStIOMap_UwRw_FE^.o_xCutHolder_DnCut					; (* 下裁刀架 *)
			o_xCutCylinder_DnCut			:= i_pstStIOMap_UwRw_FE^.o_xCutCylinder_DnCut				; (* 下裁胶辊 *)
			o_xCutter_DnCut					:= i_pstStIOMap_UwRw_FE^.o_xCutter_DnCut						; (* 下裁裁刀 *)
			o_xLamp_PaperCoreSelect6Inch	:= i_pstStIOMap_UwRw_FE^.o_xLamp_PaperCoreSelect6Inch		;(* 6寸纸管指示 *)
			o_xLamp_InverterError			:= i_pstStIOMap_UwRw_FE^.o_xLamp_InverterError				; (* 变频故障 *)
			o_xAxisATorqueCancel			:= i_pstStIOMap_UwRw_FE^.o_xAxisATorqueCancel				; (* A轴转矩取消 *)
			o_xAxisBTorqueCancel			:= i_pstStIOMap_UwRw_FE^.o_xAxisBTorqueCancel				; (* B轴转矩取消 *)
			o_wAxisATorqueVolt				:= i_pstStIOMap_UwRw_FE^.o_wAxisATorqueVolt					; (* A轴转矩电压 *)
			o_wAxisBTorqueVolt				:= i_pstStIOMap_UwRw_FE^.o_wAxisBTorqueVolt					; (* B轴转矩电压 *)
			o_xLampAxisInching				:= i_pstStIOMap_UwRw_FE^.o_xLampAxisInching					; (* 轴单运行指示 *)
			(*2024.09.28.094834//增加秦华IO*)
			o_xHydrPumpPower				:= i_pstStIOMap_UwRw_FE^.o_xHydrPumpPower					; (* 液压泵
源开关 *)
			o_xAdvanceAllBoot				:= i_pstStIOMap_UwRw_FE^.o_xAdvanceAllBoot					; (* 开机整体进版信号 *)
			o_xStopBack						:= i_pstStIOMap_UwRw_FE^.o_xStopBack							; (* 停止退版信号 *)
			//2026.05.26.145044+使用的o_xOutputAlarm未被赋值
			i_pstStIOMap_UwRw_FE^.o_xOutputAlarm:= i_pstStIOMap_UwRw_FE^.o_xRel_AlarmBell						; (* 警报输出 *)

			o_xOutputAlarm					:= i_pstStIOMap_UwRw_FE^.o_xOutputAlarm						; (* 警报输出 *)
			o_xServoError					:= i_pstStIOMap_UwRw_FE^.o_xServoError						; (* 伺服故障信号 *)

			o_xRsvd_DO0						:= i_pstStIOMap_UwRw_FE^.o_xRsvd_DO0							; (* 数字量输出保留0 *)//放卷变频器运行
			o_xRsvd_DO1						:= i_pstStIOMap_UwRw_FE^.o_xRsvd_DO1							; (* 数字量输出保留1 *)
			o_xRsvd_DO2						:= i_pstStIOMap_UwRw_FE^.o_xRsvd_DO2							; (* 数字量输出保留2 *)
			o_xRsvd_DO3						:= i_pstStIOMap_UwRw_FE^.o_xRsvd_DO3							; (* 数字量输出保留3 *)
			o_xRsvd_DO4						:= i_pstStIOMap_UwRw_FE^.o_xRsvd_DO4							; (* 数字量输出保留4 *)
			o_xRsvd_DO5						:= i_pstStIOMap_UwRw_FE^.o_xRsvd_DO5							; (* 数字量输出保留5 *)
			o_xRsvd_DO6						:= i_pstStIOMap_UwRw_FE^.o_xRsvd_DO6							; (* 数字量输出保留6 *)
			o_xRsvd_DO7						:= i_pstStIOMap_UwRw_FE^.o_xRsvd_DO7							; (* 数字量输出保留7 *)
			o_xRsvd_DO8						:= i_pstStIOMap_UwRw_FE^.o_xRsvd_DO8							; (* 数字量输出保留8 *)
			o_xRsvd_DO9						:= i_pstStIOMap_UwRw_FE^.o_xRsvd_DO9							; (* 数字量输出保留9 *)
			o_wRsvd_AO0						:= i_pstStIOMap_UwRw_FE^.o_wRsvd_AO0							; (* 模拟量输出保留0 *)//UV启动器
			o_wRsvd_AO1						:= i_pstStIOMap_UwRw_FE^.o_wRsvd_AO1							; (* 模拟量输出保留1 *)
			o_wRsvd_AO2						:= i_pstStIOMap_UwRw_FE^.o_wRsvd_AO2							; (* 模拟量输出保留2 *)
			o_wRsvd_AO3						:= i_pstStIOMap_UwRw_FE^.o_wRsvd_AO3							; (* 模拟量输出保留3 *)
			o_wRsvd_AO4						:= i_pstStIOMap_UwRw_FE^.o_wRsvd_AO4							; (* 模拟量输出保留4 *)
			o_wRsvd_AO5						:= i_pstStIOMap_UwRw_FE^.o_wRsvd_AO5							; (* 模拟量输出保留5 *)
		END_IF
	ELSE
		o_iErNo:= -1;
	END_IF
ELSE
	o_xEstopLamp					:= FALSE; (* 急停指示 *)
	o_xLamp_PreDrive				:= FALSE; (* 预驱同步指示 *)
	o_xRel_TowerForeward			:= FALSE; (* 塔台正转 *)
	o_xRel_TowerReversal			:= FALSE; (* 塔台反转 *)
	o_xAxisALamp					:= FALSE; (* A轴指示 *)
	o_xAxisBLamp					:= FALSE; (* B轴指示 *)
	o_xCutHolder_UpCut				:= FALSE; (* 上裁刀架 *)
	o_xCutCylinder_UpCut			:= FALSE; (* 上裁胶辊 *)
	o_xCutter_UpCut					:= FALSE; (* 上裁裁刀 *)
	o_xCutHolder_DnCut				:= FALSE; (* 下裁刀架 *)
	o_xCutCylinder_DnCut			:= FALSE; (* 下裁胶辊 *)
	o_xCutter_DnCut					:= FALSE; (* 下裁裁刀 *)
	o_xLamp_PaperCoreSelect6Inch	:= FALSE;(* 6寸纸管指示 *)

	o_xRsvd_DO0						:= FALSE; (* 数字量输出保留0 *)
	o_xRsvd_DO1						:= FALSE; (* 数字量输出保留1 *)
	o_xRsvd_DO2						:= FALSE; (* 数字量输出保留2 *)
	o_xRsvd_DO3						:= FALSE; (* 数字量输出保留3 *)
	o_xRsvd_DO4						:= FALSE; (* 数字量输出保留4 *)
	o_xRsvd_DO5						:= FALSE; (* 数字量输出保留5 *)
	o_xRsvd_DO6						:= FALSE; (* 数字量输出保留6 *)
	o_xRsvd_DO7						:= FALSE; (* 数字量输出保留7 *)
	o_xRsvd_DO8						:= FALSE; (* 数字量输出保留8 *)
	o_xRsvd_DO9						:= FALSE; (* 数字量输出保留9 *)
	o_wRsvd_AO0						:= 0; (* 模拟量输出保留0 *)
	o_wRsvd_AO1						:= 0; (* 模拟量输出保留1 *)
	o_wRsvd_AO2						:= 0; (* 模拟量输出保留2 *)
	o_wRsvd_AO3						:= 0; (* 模拟量输出保留3 *)
	o_wRsvd_AO4						:= 0; (* 模拟量输出保留4 *)
	o_wRsvd_AO5						:= 0; (* 模拟量输出保留5 *)
END_IF
